(* IEC 61131-3 sources: plc-st-coding-agent/progress/evidence/f14_v10_full_20261113/jobs/custom_deepseek-v4pro, 130 files *)

(* ---- public-easy-01.candidate_01.st ---- *)
(*
ENGINEERING_CONTRACT
- Pump_Motor: active in state Cleaning, set by bottleSensor true when idle, retained until cleaningConfirmButton true (PUB001-PUB003).
- Filling_Valve: active in state Filling, set by cleaningConfirmButton true in Cleaning, retained until fillingConfirmButton true (PUB003-PUB004).
- Capping_Machine: active in state Capping, set by fillingConfirmButton true in Filling, retained until cappingConfirmButton true (PUB004-PUB005).
- Packing_Machine: active in state Packing, set by cappingConfirmButton true in Capping, retained until packingConfirmButton true (PUB005-PUB006).
- Completion_Light: active in state Done, set by packingConfirmButton true in Packing, retained until finishedButton true (PUB006-PUB007).
- Same-scan priority: exactly one transition evaluated per scan via IF/ELSIF on current state; outputs updated after transition.
- Units/boundaries: all signals are BOOL; state is an integer constant 0..5; no timing or analog units involved.
*)
(* CONTRACT_RULES [] *)

FUNCTION_BLOCK AutomatedFillingLineControl
VAR CONSTANT
    ST_IDLE : INT := 0;
    ST_CLEANING : INT := 1;
    ST_FILLING : INT := 2;
    ST_CAPPING : INT := 3;
    ST_PACKING : INT := 4;
    ST_DONE : INT := 5;
END_VAR
VAR
    state : INT := 0; (* initial idle state *)
END_VAR

IF state = ST_IDLE THEN
    IF bottleSensor THEN
        state := ST_CLEANING;
    END_IF;
ELSIF state = ST_CLEANING THEN
    IF cleaningConfirmButton THEN
        state := ST_FILLING;
    END_IF;
ELSIF state = ST_FILLING THEN
    IF fillingConfirmButton THEN
        state := ST_CAPPING;
    END_IF;
ELSIF state = ST_CAPPING THEN
    IF cappingConfirmButton THEN
        state := ST_PACKING;
    END_IF;
ELSIF state = ST_PACKING THEN
    IF packingConfirmButton THEN
        state := ST_DONE;
    END_IF;
ELSIF state = ST_DONE THEN
    IF finishedButton THEN
        state := ST_IDLE;
    END_IF;
END_IF;

Pump_Motor := (state = ST_CLEANING);
Filling_Valve := (state = ST_FILLING);
Capping_Machine := (state = ST_CAPPING);
Packing_Machine := (state = ST_PACKING);
Completion_Light := (state = ST_DONE);

END_FUNCTION_BLOCK

(* ---- public-easy-01.candidate_02.st ---- *)
(*
ENGINEERING_CONTRACT
- Pump_Motor: active in state Cleaning, set by bottleSensor true when idle, retained until cleaningConfirmButton true (PUB001-PUB003).
- Filling_Valve: active in state Filling, set by cleaningConfirmButton true in Cleaning, retained until fillingConfirmButton true (PUB003-PUB004).
- Capping_Machine: active in state Capping, set by fillingConfirmButton true in Filling, retained until cappingConfirmButton true (PUB004-PUB005).
- Packing_Machine: active in state Packing, set by cappingConfirmButton true in Capping, retained until packingConfirmButton true (PUB005-PUB006).
- Completion_Light: active in state Done, set by packingConfirmButton true in Packing, retained until finishedButton true (PUB006-PUB007).
- Same-scan priority: exactly one transition evaluated per scan via IF/ELSIF on current state; outputs updated after transition.
- Units/boundaries: all signals are BOOL; state is an integer constant 0..5; no timing or analog units involved.
*)
(* CONTRACT_RULES [] *)

FUNCTION_BLOCK AutomatedFillingLineControl
VAR_INPUT
    bottleSensor : BOOL;
    cleaningConfirmButton : BOOL;
    fillingConfirmButton : BOOL;
    cappingConfirmButton : BOOL;
    packingConfirmButton : BOOL;
    finishedButton : BOOL;
END_VAR
VAR_OUTPUT
    Pump_Motor : BOOL;
    Filling_Valve : BOOL;
    Capping_Machine : BOOL;
    Packing_Machine : BOOL;
    Completion_Light : BOOL;
END_VAR
VAR CONSTANT
    ST_IDLE : INT := 0;
    ST_CLEANING : INT := 1;
    ST_FILLING : INT := 2;
    ST_CAPPING : INT := 3;
    ST_PACKING : INT := 4;
    ST_DONE : INT := 5;
END_VAR
VAR
    state : INT := 0; (* initial idle state *)
END_VAR

IF state = ST_IDLE THEN
    IF bottleSensor THEN
        state := ST_CLEANING;
    END_IF;
ELSIF state = ST_CLEANING THEN
    IF cleaningConfirmButton THEN
        state := ST_FILLING;
    END_IF;
ELSIF state = ST_FILLING THEN
    IF fillingConfirmButton THEN
        state := ST_CAPPING;
    END_IF;
ELSIF state = ST_CAPPING THEN
    IF cappingConfirmButton THEN
        state := ST_PACKING;
    END_IF;
ELSIF state = ST_PACKING THEN
    IF packingConfirmButton THEN
        state := ST_DONE;
    END_IF;
ELSIF state = ST_DONE THEN
    IF finishedButton THEN
        state := ST_IDLE;
    END_IF;
END_IF;

Pump_Motor := (state = ST_CLEANING);
Filling_Valve := (state = ST_FILLING);
Capping_Machine := (state = ST_CAPPING);
Packing_Machine := (state = ST_PACKING);
Completion_Light := (state = ST_DONE);

END_FUNCTION_BLOCK

(* ---- public-easy-01.raw_candidate_01.st ---- *)
(*
ENGINEERING_CONTRACT
- Pump_Motor: active in state Cleaning, set by bottleSensor true when idle, retained until cleaningConfirmButton true (PUB001-PUB003).
- Filling_Valve: active in state Filling, set by cleaningConfirmButton true in Cleaning, retained until fillingConfirmButton true (PUB003-PUB004).
- Capping_Machine: active in state Capping, set by fillingConfirmButton true in Filling, retained until cappingConfirmButton true (PUB004-PUB005).
- Packing_Machine: active in state Packing, set by cappingConfirmButton true in Capping, retained until packingConfirmButton true (PUB005-PUB006).
- Completion_Light: active in state Done, set by packingConfirmButton true in Packing, retained until finishedButton true (PUB006-PUB007).
- Same-scan priority: exactly one transition evaluated per scan via IF/ELSIF on current state; outputs updated after transition.
- Units/boundaries: all signals are BOOL; state is an integer constant 0..5; no timing or analog units involved.
*)
(* CONTRACT_RULES [] *)

FUNCTION_BLOCK AutomatedFillingLineControl
VAR CONSTANT
    ST_IDLE : INT := 0;
    ST_CLEANING : INT := 1;
    ST_FILLING : INT := 2;
    ST_CAPPING : INT := 3;
    ST_PACKING : INT := 4;
    ST_DONE : INT := 5;
END_VAR
VAR
    state : INT := 0; (* initial idle state *)
END_VAR

IF state = ST_IDLE THEN
    IF bottleSensor THEN
        state := ST_CLEANING;
    END_IF;
ELSIF state = ST_CLEANING THEN
    IF cleaningConfirmButton THEN
        state := ST_FILLING;
    END_IF;
ELSIF state = ST_FILLING THEN
    IF fillingConfirmButton THEN
        state := ST_CAPPING;
    END_IF;
ELSIF state = ST_CAPPING THEN
    IF cappingConfirmButton THEN
        state := ST_PACKING;
    END_IF;
ELSIF state = ST_PACKING THEN
    IF packingConfirmButton THEN
        state := ST_DONE;
    END_IF;
ELSIF state = ST_DONE THEN
    IF finishedButton THEN
        state := ST_IDLE;
    END_IF;
END_IF;

Pump_Motor := (state = ST_CLEANING);
Filling_Valve := (state = ST_FILLING);
Capping_Machine := (state = ST_CAPPING);
Packing_Machine := (state = ST_PACKING);
Completion_Light := (state = ST_DONE);

END_FUNCTION_BLOCK

(* ---- public-easy-01.raw_candidate_02.st ---- *)
(*
ENGINEERING_CONTRACT
- Pump_Motor: active in state Cleaning, set by bottleSensor true when idle, retained until cleaningConfirmButton true (PUB001-PUB003).
- Filling_Valve: active in state Filling, set by cleaningConfirmButton true in Cleaning, retained until fillingConfirmButton true (PUB003-PUB004).
- Capping_Machine: active in state Capping, set by fillingConfirmButton true in Filling, retained until cappingConfirmButton true (PUB004-PUB005).
- Packing_Machine: active in state Packing, set by cappingConfirmButton true in Capping, retained until packingConfirmButton true (PUB005-PUB006).
- Completion_Light: active in state Done, set by packingConfirmButton true in Packing, retained until finishedButton true (PUB006-PUB007).
- Same-scan priority: exactly one transition evaluated per scan via IF/ELSIF on current state; outputs updated after transition.
- Units/boundaries: all signals are BOOL; state is an integer constant 0..5; no timing or analog units involved.
*)
(* CONTRACT_RULES [] *)

FUNCTION_BLOCK AutomatedFillingLineControl
VAR_INPUT
    bottleSensor : BOOL;
    cleaningConfirmButton : BOOL;
    fillingConfirmButton : BOOL;
    cappingConfirmButton : BOOL;
    packingConfirmButton : BOOL;
    finishedButton : BOOL;
END_VAR
VAR_OUTPUT
    Pump_Motor : BOOL;
    Filling_Valve : BOOL;
    Capping_Machine : BOOL;
    Packing_Machine : BOOL;
    Completion_Light : BOOL;
END_VAR
VAR CONSTANT
    ST_IDLE : INT := 0;
    ST_CLEANING : INT := 1;
    ST_FILLING : INT := 2;
    ST_CAPPING : INT := 3;
    ST_PACKING : INT := 4;
    ST_DONE : INT := 5;
END_VAR
VAR
    state : INT := 0; (* initial idle state *)
END_VAR

IF state = ST_IDLE THEN
    IF bottleSensor THEN
        state := ST_CLEANING;
    END_IF;
ELSIF state = ST_CLEANING THEN
    IF cleaningConfirmButton THEN
        state := ST_FILLING;
    END_IF;
ELSIF state = ST_FILLING THEN
    IF fillingConfirmButton THEN
        state := ST_CAPPING;
    END_IF;
ELSIF state = ST_CAPPING THEN
    IF cappingConfirmButton THEN
        state := ST_PACKING;
    END_IF;
ELSIF state = ST_PACKING THEN
    IF packingConfirmButton THEN
        state := ST_DONE;
    END_IF;
ELSIF state = ST_DONE THEN
    IF finishedButton THEN
        state := ST_IDLE;
    END_IF;
END_IF;

Pump_Motor := (state = ST_CLEANING);
Filling_Valve := (state = ST_FILLING);
Capping_Machine := (state = ST_CAPPING);
Packing_Machine := (state = ST_PACKING);
Completion_Light := (state = ST_DONE);

END_FUNCTION_BLOCK

(* ---- public-easy-02.candidate_01.st ---- *)
(*
ENGINEERING_CONTRACT
Activation: On every call after first, edge outputs computed from value vs lastValue.
Retention/hold: No latched outputs; all outputs are recomputed each scan from current and previous DWORD.
Reset/deactivation: No explicit reset; first invocation sets baseline lastValue:=value and reports no edges.
Same-scan priority: value is captured at scan start into lastValue after output computation; simultaneous change detection only.
Units/boundaries: risingBits/fallingBits are 32-bit DWORD masks, counts 0..32 as USINT; PUB001.
*)
(* CONTRACT_RULES [] *)

FUNCTION_BLOCK FB
VAR_INPUT
    value : DWORD;
END_VAR
VAR_OUTPUT
    hasChanged : BOOL;
    hasRisingEdges : BOOL;
    risingBits : DWORD;
    noOfRisingBits : USINT;
    hasFallingEdges : BOOL;
    fallingBits : DWORD;
    noOfFallingBits : USINT;
END_VAR
VAR
    lastValue : DWORD := DWORD#0;
    initialized : BOOL := FALSE;
    tmp_bits : DWORD;
    tmp_count : USINT;
    tmp_i : USINT;
END_VAR

// On first call, initialize previous value and report no changes/edges.
IF NOT initialized THEN
    lastValue := value;
    initialized := TRUE;
    hasChanged := FALSE;
    hasRisingEdges := FALSE;
    risingBits := DWORD#0;
    noOfRisingBits := USINT#0;
    hasFallingEdges := FALSE;
    fallingBits := DWORD#0;
    noOfFallingBits := USINT#0;
    RETURN;
END_IF;

// Compute changes and edge masks.
hasChanged := (value <> lastValue);
risingBits := value AND (NOT lastValue);
fallingBits := lastValue AND (NOT value);
hasRisingEdges := (risingBits <> DWORD#0);
hasFallingEdges := (fallingBits <> DWORD#0);

// Count rising edge bits.
tmp_count := USINT#0;
tmp_bits := risingBits;
FOR tmp_i := USINT#0 TO USINT#31 DO
    IF (tmp_bits AND DWORD#1) <> DWORD#0 THEN
        tmp_count := tmp_count + USINT#1;
    END_IF;
    tmp_bits := SHR(tmp_bits, UINT#1);
END_FOR;
noOfRisingBits := tmp_count;

// Count falling edge bits.
tmp_count := USINT#0;
tmp_bits := fallingBits;
FOR tmp_i := USINT#0 TO USINT#31 DO
    IF (tmp_bits AND DWORD#1) <> DWORD#0 THEN
        tmp_count := tmp_count + USINT#1;
    END_IF;
    tmp_bits := SHR(tmp_bits, UINT#1);
END_FOR;
noOfFallingBits := tmp_count;

// Store current value for next cycle.
lastValue := value;

END_FUNCTION_BLOCK

(* ---- public-easy-02.candidate_02.st ---- *)
(*
ENGINEERING_CONTRACT
Activation: On every call including first, edge outputs computed from value versus lastValue; lastValue initializes to 0.
Retention/hold: No latched outputs; all outputs are recomputed each scan from current and previous DWORD.
Reset/deactivation: No explicit reset; first invocation compares against zero and reports rising edges for set input bits.
Same-scan priority: value is captured before output computation; lastValue is updated at the end of the same invocation.
Units/boundaries: DWORD 32-bit masks, counts 0..32 as USINT; PUB001.
*)
(* CONTRACT_RULES [] *)

FUNCTION_BLOCK FB
VAR_INPUT
    value : DWORD;
END_VAR
VAR_OUTPUT
    hasChanged : BOOL;
    hasRisingEdges : BOOL;
    risingBits : DWORD;
    noOfRisingBits : USINT;
    hasFallingEdges : BOOL;
    fallingBits : DWORD;
    noOfFallingBits : USINT;
END_VAR
VAR
    lastValue : DWORD := DWORD#0;
    tmp_bits : DWORD;
    tmp_count : USINT;
    tmp_i : USINT;
END_VAR

hasChanged := (value <> lastValue);
risingBits := value AND (NOT lastValue);
fallingBits := lastValue AND (NOT value);
hasRisingEdges := (risingBits <> DWORD#0);
hasFallingEdges := (fallingBits <> DWORD#0);

tmp_count := USINT#0;
tmp_bits := risingBits;
FOR tmp_i := USINT#0 TO USINT#31 DO
    IF (tmp_bits AND DWORD#1) <> DWORD#0 THEN
        tmp_count := tmp_count + USINT#1;
    END_IF;
    tmp_bits := SHR(tmp_bits, UINT#1);
END_FOR;
noOfRisingBits := tmp_count;

tmp_count := USINT#0;
tmp_bits := fallingBits;
FOR tmp_i := USINT#0 TO USINT#31 DO
    IF (tmp_bits AND DWORD#1) <> DWORD#0 THEN
        tmp_count := tmp_count + USINT#1;
    END_IF;
    tmp_bits := SHR(tmp_bits, UINT#1);
END_FOR;
noOfFallingBits := tmp_count;

lastValue := value;

END_FUNCTION_BLOCK

(* ---- public-easy-02.raw_candidate_01.st ---- *)
(*
ENGINEERING_CONTRACT
Activation: On every call after first, edge outputs computed from value vs lastValue.
Retention/hold: No latched outputs; all outputs are recomputed each scan from current and previous DWORD.
Reset/deactivation: No explicit reset; first invocation sets baseline lastValue:=value and reports no edges.
Same-scan priority: value is captured at scan start into lastValue after output computation; simultaneous change detection only.
Units/boundaries: risingBits/fallingBits are 32-bit DWORD masks, counts 0..32 as USINT; PUB001.
*)
(* CONTRACT_RULES [] *)

FUNCTION_BLOCK FB
VAR_INPUT
    value : DWORD;
END_VAR
VAR_OUTPUT
    hasChanged : BOOL;
    hasRisingEdges : BOOL;
    risingBits : DWORD;
    noOfRisingBits : USINT;
    hasFallingEdges : BOOL;
    fallingBits : DWORD;
    noOfFallingBits : USINT;
END_VAR
VAR
    lastValue : DWORD := DWORD#0;
    initialized : BOOL := FALSE;
    tmp_bits : DWORD;
    tmp_count : USINT;
    tmp_i : USINT;
END_VAR

// On first call, initialize previous value and report no changes/edges.
IF NOT initialized THEN
    lastValue := value;
    initialized := TRUE;
    hasChanged := FALSE;
    hasRisingEdges := FALSE;
    risingBits := DWORD#0;
    noOfRisingBits := USINT#0;
    hasFallingEdges := FALSE;
    fallingBits := DWORD#0;
    noOfFallingBits := USINT#0;
    RETURN;
END_IF;

// Compute changes and edge masks.
hasChanged := (value <> lastValue);
risingBits := value AND (NOT lastValue);
fallingBits := lastValue AND (NOT value);
hasRisingEdges := (risingBits <> DWORD#0);
hasFallingEdges := (fallingBits <> DWORD#0);

// Count rising edge bits.
tmp_count := USINT#0;
tmp_bits := risingBits;
FOR tmp_i := USINT#0 TO USINT#31 DO
    IF (tmp_bits AND DWORD#1) <> DWORD#0 THEN
        tmp_count := tmp_count + USINT#1;
    END_IF;
    tmp_bits := SHR(tmp_bits, UINT#1);
END_FOR;
noOfRisingBits := tmp_count;

// Count falling edge bits.
tmp_count := USINT#0;
tmp_bits := fallingBits;
FOR tmp_i := USINT#0 TO USINT#31 DO
    IF (tmp_bits AND DWORD#1) <> DWORD#0 THEN
        tmp_count := tmp_count + USINT#1;
    END_IF;
    tmp_bits := SHR(tmp_bits, UINT#1);
END_FOR;
noOfFallingBits := tmp_count;

// Store current value for next cycle.
lastValue := value;

END_FUNCTION_BLOCK

(* ---- public-easy-02.raw_candidate_02.st ---- *)
(*
ENGINEERING_CONTRACT
Activation: On every call including first, edge outputs computed from value versus lastValue; lastValue initializes to 0.
Retention/hold: No latched outputs; all outputs are recomputed each scan from current and previous DWORD.
Reset/deactivation: No explicit reset; first invocation compares against zero and reports rising edges for set input bits.
Same-scan priority: value is captured before output computation; lastValue is updated at the end of the same invocation.
Units/boundaries: DWORD 32-bit masks, counts 0..32 as USINT; PUB001.
*)
(* CONTRACT_RULES [] *)

FUNCTION_BLOCK FB
VAR_INPUT
    value : DWORD;
END_VAR
VAR_OUTPUT
    hasChanged : BOOL;
    hasRisingEdges : BOOL;
    risingBits : DWORD;
    noOfRisingBits : USINT;
    hasFallingEdges : BOOL;
    fallingBits : DWORD;
    noOfFallingBits : USINT;
END_VAR
VAR
    lastValue : DWORD := DWORD#0;
    tmp_bits : DWORD;
    tmp_count : USINT;
    tmp_i : USINT;
END_VAR

hasChanged := (value <> lastValue);
risingBits := value AND (NOT lastValue);
fallingBits := lastValue AND (NOT value);
hasRisingEdges := (risingBits <> DWORD#0);
hasFallingEdges := (fallingBits <> DWORD#0);

tmp_count := USINT#0;
tmp_bits := risingBits;
FOR tmp_i := USINT#0 TO USINT#31 DO
    IF (tmp_bits AND DWORD#1) <> DWORD#0 THEN
        tmp_count := tmp_count + USINT#1;
    END_IF;
    tmp_bits := SHR(tmp_bits, UINT#1);
END_FOR;
noOfRisingBits := tmp_count;

tmp_count := USINT#0;
tmp_bits := fallingBits;
FOR tmp_i := USINT#0 TO USINT#31 DO
    IF (tmp_bits AND DWORD#1) <> DWORD#0 THEN
        tmp_count := tmp_count + USINT#1;
    END_IF;
    tmp_bits := SHR(tmp_bits, UINT#1);
END_FOR;
noOfFallingBits := tmp_count;

lastValue := value;

END_FUNCTION_BLOCK

(* ---- public-easy-03.candidate_01.st ---- *)
(* ENGINEERING_CONTRACT
   hiAlarm : SET on Value > hiLevel (PUB001), RESET on Value < hiLevel-hystWindow (PUB002), otherwise hold previous state.
   loAlarm : SET on Value < loLevel (PUB003), RESET on Value > loLevel+hystWindow (PUB004), otherwise hold previous state.
   error/status : SET 16#8001 when loLevel>=hiLevel and return (PUB005); SET 16#8002 when hystWindow>=hiLevel-loLevel and return (PUB006); cleared to FALSE/0 before checks.
   Priority : error checks run before alarm update; error returns preserve last alarm outputs.
   Boundaries : strict > and < for activation/deactivation; exact threshold equality holds current state. Negative hystWindow unspecified; applied as supplied.
   Units : REAL thresholds and values; status is WORD hex code.
*)
(* CONTRACT_RULES [] *)
FUNCTION_BLOCK AlarmHandling
VAR_INPUT
    Value : REAL;
    hiLevel : REAL;
    loLevel : REAL;
    hystWindow : REAL;
END_VAR
VAR_OUTPUT
    hiAlarm : BOOL;
    loAlarm : BOOL;
    error : BOOL;
    status : WORD;
END_VAR
VAR
END_VAR

    error := FALSE;
    status := 0;

    IF loLevel >= hiLevel THEN
        error := TRUE;
        status := 16#8001;
        RETURN;
    END_IF;

    IF hystWindow >= (hiLevel - loLevel) THEN
        error := TRUE;
        status := 16#8002;
        RETURN;
    END_IF;

    IF Value > hiLevel THEN
        hiAlarm := TRUE;
    ELSIF Value < (hiLevel - hystWindow) THEN
        hiAlarm := FALSE;
    END_IF;

    IF Value < loLevel THEN
        loAlarm := TRUE;
    ELSIF Value > (loLevel + hystWindow) THEN
        loAlarm := FALSE;
    END_IF;

END_FUNCTION_BLOCK

(* ---- public-easy-03.raw_candidate_01.st ---- *)
(* ENGINEERING_CONTRACT
   hiAlarm : SET on Value > hiLevel (PUB001), RESET on Value < hiLevel-hystWindow (PUB002), otherwise hold previous state.
   loAlarm : SET on Value < loLevel (PUB003), RESET on Value > loLevel+hystWindow (PUB004), otherwise hold previous state.
   error/status : SET 16#8001 when loLevel>=hiLevel and return (PUB005); SET 16#8002 when hystWindow>=hiLevel-loLevel and return (PUB006); cleared to FALSE/0 before checks.
   Priority : error checks run before alarm update; error returns preserve last alarm outputs.
   Boundaries : strict > and < for activation/deactivation; exact threshold equality holds current state. Negative hystWindow unspecified; applied as supplied.
   Units : REAL thresholds and values; status is WORD hex code.
*)
(* CONTRACT_RULES [] *)
FUNCTION_BLOCK AlarmHandling
VAR_INPUT
    Value : REAL;
    hiLevel : REAL;
    loLevel : REAL;
    hystWindow : REAL;
END_VAR
VAR_OUTPUT
    hiAlarm : BOOL;
    loAlarm : BOOL;
    error : BOOL;
    status : WORD;
END_VAR
VAR
END_VAR

    error := FALSE;
    status := 0;

    IF loLevel >= hiLevel THEN
        error := TRUE;
        status := 16#8001;
        RETURN;
    END_IF;

    IF hystWindow >= (hiLevel - loLevel) THEN
        error := TRUE;
        status := 16#8002;
        RETURN;
    END_IF;

    IF Value > hiLevel THEN
        hiAlarm := TRUE;
    ELSIF Value < (hiLevel - hystWindow) THEN
        hiAlarm := FALSE;
    END_IF;

    IF Value < loLevel THEN
        loAlarm := TRUE;
    ELSIF Value > (loLevel + hystWindow) THEN
        loAlarm := FALSE;
    END_IF;

END_FUNCTION_BLOCK

(* ---- public-easy-04.candidate_01.st ---- *)
(*
ENGINEERING_CONTRACT
1. DebounceValid state: set only while VISCOSITY_OK=TRUE and PASTE_E_STOP_NC=TRUE after accumulated CycleTime >= DebounceTime; immediate invalidation when VISCOSITY_OK=FALSE; incomplete timing is cleared when E-stop is FALSE (PUB001, PUB002).
2. VFD_RUN: active = PASTE_E_STOP_NC AND DebounceValid; E-stop has immediate priority and disables output in the same scan; no output latching (PUB002).
3. PUMP_RUNTIME_ACC: accumulates TO_LTIME(CycleTime) only when same-scan VFD_RUN=TRUE; preserves accumulated time while stopped; initial value 0 (PUB003, PUB005).
4. PUMP_MAINT_DUE: set when PUMP_RUNTIME_ACC >= LTIME#500H; because runtime is monotonic, it remains set; informational only with no effect on run/permissive logic (PUB004).
5. Initialization: VFD_RUN=FALSE, PUMP_RUNTIME_ACC=LTIME#0S, PUMP_MAINT_DUE=FALSE via declared initial values (PUB005).
Boundary: threshold comparisons use >= and TIME values are converted to LTIME; first satisfying debounce tick occurs when accumulated CycleTime reaches DebounceTime.
Unspecified: non-positive DebounceTime or CycleTime are assumed to be supplied positive (PUB006).
*)
(* CONTRACT_RULES [] *)
FUNCTION_BLOCK JamPump
VAR_INPUT
    VISCOSITY_OK : BOOL;
    PASTE_E_STOP_NC : BOOL;
    DebounceTime : TIME;
    CycleTime : TIME;
END_VAR
VAR_OUTPUT
    VFD_RUN : BOOL := FALSE;
    PUMP_MAINT_DUE : BOOL := FALSE;
    PUMP_RUNTIME_ACC : LTIME := LTIME#0S;
END_VAR
VAR
    local_DebounceElapsed : LTIME := LTIME#0S;
    local_ViscCondValid : BOOL := FALSE;
    local_MaintenanceLimit : LTIME := LTIME#500H;
END_VAR

IF NOT VISCOSITY_OK THEN
    local_ViscCondValid := FALSE;
    local_DebounceElapsed := LTIME#0S;
ELSE
    IF NOT PASTE_E_STOP_NC THEN
        IF NOT local_ViscCondValid THEN
            local_DebounceElapsed := LTIME#0S;
        END_IF;
    ELSE
        IF NOT local_ViscCondValid THEN
            local_DebounceElapsed := local_DebounceElapsed + TO_LTIME(CycleTime);
            IF local_DebounceElapsed >= TO_LTIME(DebounceTime) THEN
                local_ViscCondValid := TRUE;
            END_IF;
        END_IF;
    END_IF;
END_IF;

VFD_RUN := PASTE_E_STOP_NC AND local_ViscCondValid;

IF VFD_RUN THEN
    PUMP_RUNTIME_ACC := PUMP_RUNTIME_ACC + TO_LTIME(CycleTime);
END_IF;

PUMP_MAINT_DUE := (PUMP_RUNTIME_ACC >= local_MaintenanceLimit);

END_FUNCTION_BLOCK

(* ---- public-easy-04.raw_candidate_01.st ---- *)
(*
ENGINEERING_CONTRACT
1. DebounceValid state: set only while VISCOSITY_OK=TRUE and PASTE_E_STOP_NC=TRUE after accumulated CycleTime >= DebounceTime; immediate invalidation when VISCOSITY_OK=FALSE; incomplete timing is cleared when E-stop is FALSE (PUB001, PUB002).
2. VFD_RUN: active = PASTE_E_STOP_NC AND DebounceValid; E-stop has immediate priority and disables output in the same scan; no output latching (PUB002).
3. PUMP_RUNTIME_ACC: accumulates TO_LTIME(CycleTime) only when same-scan VFD_RUN=TRUE; preserves accumulated time while stopped; initial value 0 (PUB003, PUB005).
4. PUMP_MAINT_DUE: set when PUMP_RUNTIME_ACC >= LTIME#500H; because runtime is monotonic, it remains set; informational only with no effect on run/permissive logic (PUB004).
5. Initialization: VFD_RUN=FALSE, PUMP_RUNTIME_ACC=LTIME#0S, PUMP_MAINT_DUE=FALSE via declared initial values (PUB005).
Boundary: threshold comparisons use >= and TIME values are converted to LTIME; first satisfying debounce tick occurs when accumulated CycleTime reaches DebounceTime.
Unspecified: non-positive DebounceTime or CycleTime are assumed to be supplied positive (PUB006).
*)
(* CONTRACT_RULES [] *)
FUNCTION_BLOCK JamPump
VAR_INPUT
    VISCOSITY_OK : BOOL;
    PASTE_E_STOP_NC : BOOL;
    DebounceTime : TIME;
    CycleTime : TIME;
END_VAR
VAR_OUTPUT
    VFD_RUN : BOOL := FALSE;
    PUMP_MAINT_DUE : BOOL := FALSE;
    PUMP_RUNTIME_ACC : LTIME := LTIME#0S;
END_VAR
VAR
    local_DebounceElapsed : LTIME := LTIME#0S;
    local_ViscCondValid : BOOL := FALSE;
    local_MaintenanceLimit : LTIME := LTIME#500H;
END_VAR

IF NOT VISCOSITY_OK THEN
    local_ViscCondValid := FALSE;
    local_DebounceElapsed := LTIME#0S;
ELSE
    IF NOT PASTE_E_STOP_NC THEN
        IF NOT local_ViscCondValid THEN
            local_DebounceElapsed := LTIME#0S;
        END_IF;
    ELSE
        IF NOT local_ViscCondValid THEN
            local_DebounceElapsed := local_DebounceElapsed + TO_LTIME(CycleTime);
            IF local_DebounceElapsed >= TO_LTIME(DebounceTime) THEN
                local_ViscCondValid := TRUE;
            END_IF;
        END_IF;
    END_IF;
END_IF;

VFD_RUN := PASTE_E_STOP_NC AND local_ViscCondValid;

IF VFD_RUN THEN
    PUMP_RUNTIME_ACC := PUMP_RUNTIME_ACC + TO_LTIME(CycleTime);
END_IF;

PUMP_MAINT_DUE := (PUMP_RUNTIME_ACC >= local_MaintenanceLimit);

END_FUNCTION_BLOCK

(* ---- public-easy-05.candidate_01.st ---- *)
FUNCTION_BLOCK WeldGapAlarm
VAR_INPUT
    Gap_Exceeded: BOOL;
    Weld_E_Stop_NC: BOOL;
    DebounceTime: TIME;
END_VAR
VAR_OUTPUT
    Operator_Alert: BOOL;
    Weld_Soft_Start_Active: BOOL;
END_VAR
VAR
    tmp_InitTimer: TON;
    tmp_DebounceTimer: TON;
    local_InitActive: BOOL;
    local_EStopActive: BOOL;
    local_DebounceEnable: BOOL;
END_VAR

(* ENGINEERING_CONTRACT
   Output/Group         Activation                                      Retention/Hold                     Explicit Reset/Deactivation       Same-scan priority        Units/Bounds                  PUB
   Operator_Alert       Gap_Exceeded TRUE for DebounceTime after init   Holds while eligible gap TRUE      Gap FALSE, E-stop FALSE, init   E-stop overrides monitor   TIME, positive assumed        PUB003 PUB004
   Weld_Soft_Start_Act  5 s power-up init timer not elapsed             TRUE during init unless E-stop    E-stop active, timer elapsed     E-stop overrides init       TIME 5 s                      PUB002 PUB004 PUB005
   Debounce timing      eligible gap TRUE in normal monitoring         accumulates only if eligible       Gap FALSE, E-stop, init         E-stop/init clear timing    DebounceTime TIME             PUB002 PUB003 PUB004
*)

(* CONTRACT_RULES [] *)

local_EStopActive := NOT Weld_E_Stop_NC;

tmp_InitTimer(IN := TRUE, PT := T#5S);
local_InitActive := NOT tmp_InitTimer.Q;

local_DebounceEnable := Gap_Exceeded AND NOT local_InitActive AND NOT local_EStopActive;
tmp_DebounceTimer(IN := local_DebounceEnable, PT := DebounceTime);

Operator_Alert := tmp_DebounceTimer.Q AND NOT local_EStopActive;
Weld_Soft_Start_Active := local_InitActive AND NOT local_EStopActive;

END_FUNCTION_BLOCK

(* ---- public-easy-05.raw_candidate_01.st ---- *)
FUNCTION_BLOCK WeldGapAlarm
VAR_INPUT
    Gap_Exceeded: BOOL;
    Weld_E_Stop_NC: BOOL;
    DebounceTime: TIME;
END_VAR
VAR_OUTPUT
    Operator_Alert: BOOL;
    Weld_Soft_Start_Active: BOOL;
END_VAR
VAR
    tmp_InitTimer: TON;
    tmp_DebounceTimer: TON;
    local_InitActive: BOOL;
    local_EStopActive: BOOL;
    local_DebounceEnable: BOOL;
END_VAR

(* ENGINEERING_CONTRACT
   Output/Group         Activation                                      Retention/Hold                     Explicit Reset/Deactivation       Same-scan priority        Units/Bounds                  PUB
   Operator_Alert       Gap_Exceeded TRUE for DebounceTime after init   Holds while eligible gap TRUE      Gap FALSE, E-stop FALSE, init   E-stop overrides monitor   TIME, positive assumed        PUB003 PUB004
   Weld_Soft_Start_Act  5 s power-up init timer not elapsed             TRUE during init unless E-stop    E-stop active, timer elapsed     E-stop overrides init       TIME 5 s                      PUB002 PUB004 PUB005
   Debounce timing      eligible gap TRUE in normal monitoring         accumulates only if eligible       Gap FALSE, E-stop, init         E-stop/init clear timing    DebounceTime TIME             PUB002 PUB003 PUB004
*)

(* CONTRACT_RULES [] *)

local_EStopActive := NOT Weld_E_Stop_NC;

tmp_InitTimer(IN := TRUE, PT := T#5S);
local_InitActive := NOT tmp_InitTimer.Q;

local_DebounceEnable := Gap_Exceeded AND NOT local_InitActive AND NOT local_EStopActive;
tmp_DebounceTimer(IN := local_DebounceEnable, PT := DebounceTime);

Operator_Alert := tmp_DebounceTimer.Q AND NOT local_EStopActive;
Weld_Soft_Start_Active := local_InitActive AND NOT local_EStopActive;

END_FUNCTION_BLOCK

(* ---- public-easy-06.candidate_01.st ---- *)
FUNCTION_BLOCK AerationBlowerDelayedStart
VAR_INPUT
    DO_LOW : BOOL;
    AERATION_E_STOP_NC : BOOL;
END_VAR
VAR_OUTPUT
    BLOWER_RUN : BOOL := FALSE;
    AERATION_BLOWER_CYCLE_COUNT : UINT := 0;
END_VAR
VAR
    startTimer : TON;
    startEdge : R_TRIG;
END_VAR

(*
ENGINEERING_CONTRACT
Output BLOWER_RUN:
  activation: startTimer.Q after DO_LOW AND AERATION_E_STOP_NC true for T#5S (PUB001).
  hold: remains TRUE while both inputs stay TRUE (PUB001).
  reset/deactivation: DO_LOW=FALSE or AERATION_E_STOP_NC=FALSE disables same scan and resets timer (PUB002).
  units/boundaries: BOOL.
Output AERATION_BLOWER_CYCLE_COUNT:
  activation: increment on R_TRIG false->true of BLOWER_RUN (PUB003).
  hold: retains value during operation; stop does not reset count.
  reset: only power-up/cold init to 0 (PUB004).
  units/boundaries: UINT starts; saturates at 65535 (unspecified).
*)

(* CONTRACT_RULES [] *)

startTimer(IN := DO_LOW AND AERATION_E_STOP_NC, PT := T#5S);
BLOWER_RUN := startTimer.Q;

startEdge(CLK := BLOWER_RUN);
IF startEdge.Q THEN
    IF AERATION_BLOWER_CYCLE_COUNT < UINT#65535 THEN
        AERATION_BLOWER_CYCLE_COUNT := AERATION_BLOWER_CYCLE_COUNT + UINT#1;
    END_IF;
END_IF;

END_FUNCTION_BLOCK

(* ---- public-easy-06.raw_candidate_01.st ---- *)
FUNCTION_BLOCK AerationBlowerDelayedStart
VAR_INPUT
    DO_LOW : BOOL;
    AERATION_E_STOP_NC : BOOL;
END_VAR
VAR_OUTPUT
    BLOWER_RUN : BOOL := FALSE;
    AERATION_BLOWER_CYCLE_COUNT : UINT := 0;
END_VAR
VAR
    startTimer : TON;
    startEdge : R_TRIG;
END_VAR

(*
ENGINEERING_CONTRACT
Output BLOWER_RUN:
  activation: startTimer.Q after DO_LOW AND AERATION_E_STOP_NC true for T#5S (PUB001).
  hold: remains TRUE while both inputs stay TRUE (PUB001).
  reset/deactivation: DO_LOW=FALSE or AERATION_E_STOP_NC=FALSE disables same scan and resets timer (PUB002).
  units/boundaries: BOOL.
Output AERATION_BLOWER_CYCLE_COUNT:
  activation: increment on R_TRIG false->true of BLOWER_RUN (PUB003).
  hold: retains value during operation; stop does not reset count.
  reset: only power-up/cold init to 0 (PUB004).
  units/boundaries: UINT starts; saturates at 65535 (unspecified).
*)

(* CONTRACT_RULES [] *)

startTimer(IN := DO_LOW AND AERATION_E_STOP_NC, PT := T#5S);
BLOWER_RUN := startTimer.Q;

startEdge(CLK := BLOWER_RUN);
IF startEdge.Q THEN
    IF AERATION_BLOWER_CYCLE_COUNT < UINT#65535 THEN
        AERATION_BLOWER_CYCLE_COUNT := AERATION_BLOWER_CYCLE_COUNT + UINT#1;
    END_IF;
END_IF;

END_FUNCTION_BLOCK

(* ---- public-hard-01.candidate_01.st ---- *)
(* ENGINEERING_CONTRACT
   valveARun / valveBRun / valveCRun / valveDRun / mixMotorRun:
   - Activation: manual rising-edge toggle per PUB001; auto STATES OPEN_A/OPEN_B/WAIT_C/DONE/MIXING per PUB005-PUB010.
   - Retention: hold while selected mode/state condition remains; manual toggles hold until next edge, estop FALSE, or mode change.
   - Reset/deactivation: estop=FALSE forces all FALSE and resets manual/auto state; auto transitions close prior actuator; autoStart restart wins after transitions.
   - Same-scan priority: estop overrides all; manual outputs assigned only in manual; auto transitions selected on old state, then autoStart assignment wins.
   - levelSensor units cm, thresholds >=50, >=80, >=100; processMode sampled at 80 cm branch; mixMotorComplete edge accepted only while auto MIXING.
   - Unspecified: mode switch retains auto state; after estop clear, auto requires autoStart; manual requires button restart.
*)
(* CONTRACT_RULES [] *)

TYPE AUTO_STATE : (IDLE, OPEN_A, OPEN_B, WAIT_C, MIXING, DONE);
END_TYPE;

FUNCTION_BLOCK MaterialProportioningProcessControl
VAR_INPUT
    estop : BOOL;
    opeMode : BOOL;
    valveAStart : BOOL;
    valveBStart : BOOL;
    valveCStart : BOOL;
    valveDStart : BOOL;
    mixMotorStart : BOOL;
    autoStart : BOOL;
    processMode : BOOL;
    levelSensor : INT;
    mixMotorComplete : BOOL;
END_VAR
VAR_OUTPUT
    valveARun : BOOL;
    valveBRun : BOOL;
    valveCRun : BOOL;
    valveDRun : BOOL;
    mixMotorRun : BOOL;
END_VAR
VAR
    manualValveA : BOOL := FALSE;
    manualValveB : BOOL := FALSE;
    manualValveC : BOOL := FALSE;
    manualValveD : BOOL := FALSE;
    manualMixMotor : BOOL := FALSE;

    autoState : AUTO_STATE := AUTO_STATE#IDLE;

    rt_valveA : R_TRIG;
    rt_valveB : R_TRIG;
    rt_valveC : R_TRIG;
    rt_valveD : R_TRIG;
    rt_mixMotor : R_TRIG;
    rt_autoStart : R_TRIG;
    rt_mixComplete : R_TRIG;

    tmp_autoValveA : BOOL;
    tmp_autoValveB : BOOL;
    tmp_autoValveC : BOOL;
    tmp_autoValveD : BOOL;
    tmp_autoMixMotor : BOOL;
END_VAR

// Update rising-edge detectors
rt_valveA(CLK := valveAStart);
rt_valveB(CLK := valveBStart);
rt_valveC(CLK := valveCStart);
rt_valveD(CLK := valveDStart);
rt_mixMotor(CLK := mixMotorStart);
rt_autoStart(CLK := autoStart);
rt_mixComplete(CLK := mixMotorComplete);

// Emergency stop: reset all retained states while estop is FALSE
IF NOT estop THEN
    manualValveA := FALSE;
    manualValveB := FALSE;
    manualValveC := FALSE;
    manualValveD := FALSE;
    manualMixMotor := FALSE;
    autoState := AUTO_STATE#IDLE;
END_IF;

// Manual toggle controls only in manual mode with no emergency stop
IF estop AND NOT opeMode THEN
    IF rt_valveA.Q THEN
        manualValveA := NOT manualValveA;
    END_IF;
    IF rt_valveB.Q THEN
        manualValveB := NOT manualValveB;
    END_IF;
    IF rt_valveC.Q THEN
        manualValveC := NOT manualValveC;
    END_IF;
    IF rt_valveD.Q THEN
        manualValveD := NOT manualValveD;
    END_IF;
    IF rt_mixMotor.Q THEN
        manualMixMotor := NOT manualMixMotor;
    END_IF;
END_IF;

// Automatic process state transitions
IF estop AND opeMode THEN
    CASE autoState OF
        AUTO_STATE#OPEN_A:
            IF levelSensor >= 50 THEN
                autoState := AUTO_STATE#OPEN_B;
            END_IF;

        AUTO_STATE#OPEN_B:
            IF levelSensor >= 80 THEN
                IF NOT processMode THEN
                    autoState := AUTO_STATE#MIXING;
                ELSE
                    autoState := AUTO_STATE#WAIT_C;
                END_IF;
            END_IF;

        AUTO_STATE#WAIT_C:
            IF levelSensor >= 100 THEN
                autoState := AUTO_STATE#MIXING;
            END_IF;

        AUTO_STATE#MIXING:
            IF rt_mixComplete.Q THEN
                autoState := AUTO_STATE#DONE;
            END_IF;
    END_CASE;
END_IF;

// Auto start restarts the sequence and wins over same-scan state transitions
IF estop AND opeMode AND rt_autoStart.Q THEN
    autoState := AUTO_STATE#OPEN_A;
END_IF;

// Compute temporary automatic outputs from current state
tmp_autoValveA := FALSE;
tmp_autoValveB := FALSE;
tmp_autoValveC := FALSE;
tmp_autoValveD := FALSE;
tmp_autoMixMotor := FALSE;

CASE autoState OF
    AUTO_STATE#OPEN_A:
        tmp_autoValveA := TRUE;
    AUTO_STATE#OPEN_B:
        tmp_autoValveB := TRUE;
    AUTO_STATE#WAIT_C:
        tmp_autoValveC := TRUE;
    AUTO_STATE#MIXING:
        tmp_autoMixMotor := TRUE;
    AUTO_STATE#DONE:
        tmp_autoValveD := TRUE;
END_CASE;

// Final output assignment with emergency stop as highest priority
valveARun := FALSE;
valveBRun := FALSE;
valveCRun := FALSE;
valveDRun := FALSE;
mixMotorRun := FALSE;

IF estop AND NOT opeMode THEN
    valveARun := manualValveA;
    valveBRun := manualValveB;
    valveCRun := manualValveC;
    valveDRun := manualValveD;
    mixMotorRun := manualMixMotor;
ELSIF estop AND opeMode THEN
    valveARun := tmp_autoValveA;
    valveBRun := tmp_autoValveB;
    valveCRun := tmp_autoValveC;
    valveDRun := tmp_autoValveD;
    mixMotorRun := tmp_autoMixMotor;
END_IF;

END_FUNCTION_BLOCK

(* ---- public-hard-01.candidate_02.st ---- *)
(* ENGINEERING_CONTRACT
   valveARun / valveBRun / valveCRun / valveDRun / mixMotorRun:
   - Activation: manual rising-edge toggle per PUB001; auto STATES OPEN_A/OPEN_B/WAIT_C/DONE/MIXING per PUB005-PUB010.
   - Retention: hold while selected mode/state condition remains; manual toggles hold until next edge, estop FALSE, or mode change.
   - Reset/deactivation: estop=FALSE forces all FALSE and resets manual/auto state; auto transitions close prior actuator; autoStart restart wins after transitions.
   - Same-scan priority: estop overrides all; manual outputs assigned only in manual; auto transitions selected on old state, then autoStart assignment wins.
   - levelSensor units cm, thresholds >=50, >=80, >=100; processMode sampled at 80 cm branch; mixMotorComplete edge accepted only while auto MIXING.
   - Unspecified: mode switch retains auto state; after estop clear, auto requires autoStart; manual requires button restart.
*)
(* CONTRACT_RULES [] *)

TYPE AUTO_STATE : (IDLE, OPEN_A, OPEN_B, WAIT_C, MIXING, DONE);
END_TYPE;

FUNCTION_BLOCK MaterialProportioningProcessControl
VAR_INPUT
    estop : BOOL;
    opeMode : BOOL;
    valveAStart : BOOL;
    valveBStart : BOOL;
    valveCStart : BOOL;
    valveDStart : BOOL;
    mixMotorStart : BOOL;
    autoStart : BOOL;
    processMode : BOOL;
    levelSensor : INT;
    mixMotorComplete : BOOL;
END_VAR
VAR_OUTPUT
    valveARun : BOOL;
    valveBRun : BOOL;
    valveCRun : BOOL;
    valveDRun : BOOL;
    mixMotorRun : BOOL;
END_VAR
VAR
    manualValveA : BOOL := FALSE;
    manualValveB : BOOL := FALSE;
    manualValveC : BOOL := FALSE;
    manualValveD : BOOL := FALSE;
    manualMixMotor : BOOL := FALSE;

    autoState : AUTO_STATE := IDLE;

    rt_valveA : R_TRIG;
    rt_valveB : R_TRIG;
    rt_valveC : R_TRIG;
    rt_valveD : R_TRIG;
    rt_mixMotor : R_TRIG;
    rt_autoStart : R_TRIG;
    rt_mixComplete : R_TRIG;

    tmp_autoValveA : BOOL;
    tmp_autoValveB : BOOL;
    tmp_autoValveC : BOOL;
    tmp_autoValveD : BOOL;
    tmp_autoMixMotor : BOOL;
END_VAR

// Update rising-edge detectors
rt_valveA(CLK := valveAStart);
rt_valveB(CLK := valveBStart);
rt_valveC(CLK := valveCStart);
rt_valveD(CLK := valveDStart);
rt_mixMotor(CLK := mixMotorStart);
rt_autoStart(CLK := autoStart);
rt_mixComplete(CLK := mixMotorComplete);

// Emergency stop: reset all retained states while estop is FALSE
IF NOT estop THEN
    manualValveA := FALSE;
    manualValveB := FALSE;
    manualValveC := FALSE;
    manualValveD := FALSE;
    manualMixMotor := FALSE;
    autoState := IDLE;
END_IF;

// Manual toggle controls only in manual mode with no emergency stop
IF estop AND NOT opeMode THEN
    IF rt_valveA.Q THEN
        manualValveA := NOT manualValveA;
    END_IF;
    IF rt_valveB.Q THEN
        manualValveB := NOT manualValveB;
    END_IF;
    IF rt_valveC.Q THEN
        manualValveC := NOT manualValveC;
    END_IF;
    IF rt_valveD.Q THEN
        manualValveD := NOT manualValveD;
    END_IF;
    IF rt_mixMotor.Q THEN
        manualMixMotor := NOT manualMixMotor;
    END_IF;
END_IF;

// Automatic process state transitions
IF estop AND opeMode THEN
    CASE autoState OF
        OPEN_A:
            IF levelSensor >= 50 THEN
                autoState := OPEN_B;
            END_IF;

        OPEN_B:
            IF levelSensor >= 80 THEN
                IF NOT processMode THEN
                    autoState := MIXING;
                ELSE
                    autoState := WAIT_C;
                END_IF;
            END_IF;

        WAIT_C:
            IF levelSensor >= 100 THEN
                autoState := MIXING;
            END_IF;

        MIXING:
            IF rt_mixComplete.Q THEN
                autoState := DONE;
            END_IF;
    END_CASE;
END_IF;

// Auto start restarts the sequence and wins over same-scan state transitions
IF estop AND opeMode AND rt_autoStart.Q THEN
    autoState := OPEN_A;
END_IF;

// Compute temporary automatic outputs from current state
tmp_autoValveA := FALSE;
tmp_autoValveB := FALSE;
tmp_autoValveC := FALSE;
tmp_autoValveD := FALSE;
tmp_autoMixMotor := FALSE;

CASE autoState OF
    OPEN_A:
        tmp_autoValveA := TRUE;
    OPEN_B:
        tmp_autoValveB := TRUE;
    WAIT_C:
        tmp_autoValveC := TRUE;
    MIXING:
        tmp_autoMixMotor := TRUE;
    DONE:
        tmp_autoValveD := TRUE;
END_CASE;

// Final output assignment with emergency stop as highest priority
valveARun := FALSE;
valveBRun := FALSE;
valveCRun := FALSE;
valveDRun := FALSE;
mixMotorRun := FALSE;

IF estop AND NOT opeMode THEN
    valveARun := manualValveA;
    valveBRun := manualValveB;
    valveCRun := manualValveC;
    valveDRun := manualValveD;
    mixMotorRun := manualMixMotor;
ELSIF estop AND opeMode THEN
    valveARun := tmp_autoValveA;
    valveBRun := tmp_autoValveB;
    valveCRun := tmp_autoValveC;
    valveDRun := tmp_autoValveD;
    mixMotorRun := tmp_autoMixMotor;
END_IF;

END_FUNCTION_BLOCK

(* ---- public-hard-01.raw_candidate_01.st ---- *)
(* ENGINEERING_CONTRACT
   valveARun / valveBRun / valveCRun / valveDRun / mixMotorRun:
   - Activation: manual rising-edge toggle per PUB001; auto STATES OPEN_A/OPEN_B/WAIT_C/DONE/MIXING per PUB005-PUB010.
   - Retention: hold while selected mode/state condition remains; manual toggles hold until next edge, estop FALSE, or mode change.
   - Reset/deactivation: estop=FALSE forces all FALSE and resets manual/auto state; auto transitions close prior actuator; autoStart restart wins after transitions.
   - Same-scan priority: estop overrides all; manual outputs assigned only in manual; auto transitions selected on old state, then autoStart assignment wins.
   - levelSensor units cm, thresholds >=50, >=80, >=100; processMode sampled at 80 cm branch; mixMotorComplete edge accepted only while auto MIXING.
   - Unspecified: mode switch retains auto state; after estop clear, auto requires autoStart; manual requires button restart.
*)
(* CONTRACT_RULES [] *)

TYPE AUTO_STATE : (IDLE, OPEN_A, OPEN_B, WAIT_C, MIXING, DONE);
END_TYPE

FUNCTION_BLOCK MaterialProportioningProcessControl
VAR_INPUT
    estop : BOOL;
    opeMode : BOOL;
    valveAStart : BOOL;
    valveBStart : BOOL;
    valveCStart : BOOL;
    valveDStart : BOOL;
    mixMotorStart : BOOL;
    autoStart : BOOL;
    processMode : BOOL;
    levelSensor : INT;
    mixMotorComplete : BOOL;
END_VAR
VAR_OUTPUT
    valveARun : BOOL;
    valveBRun : BOOL;
    valveCRun : BOOL;
    valveDRun : BOOL;
    mixMotorRun : BOOL;
END_VAR
VAR
    manualValveA : BOOL := FALSE;
    manualValveB : BOOL := FALSE;
    manualValveC : BOOL := FALSE;
    manualValveD : BOOL := FALSE;
    manualMixMotor : BOOL := FALSE;

    autoState : AUTO_STATE := AUTO_STATE#IDLE;

    rt_valveA : R_TRIG;
    rt_valveB : R_TRIG;
    rt_valveC : R_TRIG;
    rt_valveD : R_TRIG;
    rt_mixMotor : R_TRIG;
    rt_autoStart : R_TRIG;
    rt_mixComplete : R_TRIG;

    tmp_autoValveA : BOOL;
    tmp_autoValveB : BOOL;
    tmp_autoValveC : BOOL;
    tmp_autoValveD : BOOL;
    tmp_autoMixMotor : BOOL;
END_VAR

// Update rising-edge detectors
rt_valveA(CLK := valveAStart);
rt_valveB(CLK := valveBStart);
rt_valveC(CLK := valveCStart);
rt_valveD(CLK := valveDStart);
rt_mixMotor(CLK := mixMotorStart);
rt_autoStart(CLK := autoStart);
rt_mixComplete(CLK := mixMotorComplete);

// Emergency stop: reset all retained states while estop is FALSE
IF NOT estop THEN
    manualValveA := FALSE;
    manualValveB := FALSE;
    manualValveC := FALSE;
    manualValveD := FALSE;
    manualMixMotor := FALSE;
    autoState := AUTO_STATE#IDLE;
END_IF

// Manual toggle controls only in manual mode with no emergency stop
IF estop AND NOT opeMode THEN
    IF rt_valveA.Q THEN
        manualValveA := NOT manualValveA;
    END_IF
    IF rt_valveB.Q THEN
        manualValveB := NOT manualValveB;
    END_IF
    IF rt_valveC.Q THEN
        manualValveC := NOT manualValveC;
    END_IF
    IF rt_valveD.Q THEN
        manualValveD := NOT manualValveD;
    END_IF
    IF rt_mixMotor.Q THEN
        manualMixMotor := NOT manualMixMotor;
    END_IF
END_IF

// Automatic process state transitions
IF estop AND opeMode THEN
    CASE autoState OF
        AUTO_STATE#OPEN_A:
            IF levelSensor >= 50 THEN
                autoState := AUTO_STATE#OPEN_B;
            END_IF

        AUTO_STATE#OPEN_B:
            IF levelSensor >= 80 THEN
                IF NOT processMode THEN
                    autoState := AUTO_STATE#MIXING;
                ELSE
                    autoState := AUTO_STATE#WAIT_C;
                END_IF
            END_IF

        AUTO_STATE#WAIT_C:
            IF levelSensor >= 100 THEN
                autoState := AUTO_STATE#MIXING;
            END_IF

        AUTO_STATE#MIXING:
            IF rt_mixComplete.Q THEN
                autoState := AUTO_STATE#DONE;
            END_IF
    END_CASE
END_IF

// Auto start restarts the sequence and wins over same-scan state transitions
IF estop AND opeMode AND rt_autoStart.Q THEN
    autoState := AUTO_STATE#OPEN_A;
END_IF

// Compute temporary automatic outputs from current state
tmp_autoValveA := FALSE;
tmp_autoValveB := FALSE;
tmp_autoValveC := FALSE;
tmp_autoValveD := FALSE;
tmp_autoMixMotor := FALSE;

CASE autoState OF
    AUTO_STATE#OPEN_A:
        tmp_autoValveA := TRUE;
    AUTO_STATE#OPEN_B:
        tmp_autoValveB := TRUE;
    AUTO_STATE#WAIT_C:
        tmp_autoValveC := TRUE;
    AUTO_STATE#MIXING:
        tmp_autoMixMotor := TRUE;
    AUTO_STATE#DONE:
        tmp_autoValveD := TRUE;
END_CASE

// Final output assignment with emergency stop as highest priority
valveARun := FALSE;
valveBRun := FALSE;
valveCRun := FALSE;
valveDRun := FALSE;
mixMotorRun := FALSE;

IF estop AND NOT opeMode THEN
    valveARun := manualValveA;
    valveBRun := manualValveB;
    valveCRun := manualValveC;
    valveDRun := manualValveD;
    mixMotorRun := manualMixMotor;
ELSIF estop AND opeMode THEN
    valveARun := tmp_autoValveA;
    valveBRun := tmp_autoValveB;
    valveCRun := tmp_autoValveC;
    valveDRun := tmp_autoValveD;
    mixMotorRun := tmp_autoMixMotor;
END_IF

END_FUNCTION_BLOCK

(* ---- public-hard-01.raw_candidate_02.st ---- *)
(* ENGINEERING_CONTRACT
   valveARun / valveBRun / valveCRun / valveDRun / mixMotorRun:
   - Activation: manual rising-edge toggle per PUB001; auto STATES OPEN_A/OPEN_B/WAIT_C/DONE/MIXING per PUB005-PUB010.
   - Retention: hold while selected mode/state condition remains; manual toggles hold until next edge, estop FALSE, or mode change.
   - Reset/deactivation: estop=FALSE forces all FALSE and resets manual/auto state; auto transitions close prior actuator; autoStart restart wins after transitions.
   - Same-scan priority: estop overrides all; manual outputs assigned only in manual; auto transitions selected on old state, then autoStart assignment wins.
   - levelSensor units cm, thresholds >=50, >=80, >=100; processMode sampled at 80 cm branch; mixMotorComplete edge accepted only while auto MIXING.
   - Unspecified: mode switch retains auto state; after estop clear, auto requires autoStart; manual requires button restart.
*)
(* CONTRACT_RULES [] *)

TYPE AUTO_STATE : (IDLE, OPEN_A, OPEN_B, WAIT_C, MIXING, DONE);
END_TYPE;

FUNCTION_BLOCK MaterialProportioningProcessControl
VAR_INPUT
    estop : BOOL;
    opeMode : BOOL;
    valveAStart : BOOL;
    valveBStart : BOOL;
    valveCStart : BOOL;
    valveDStart : BOOL;
    mixMotorStart : BOOL;
    autoStart : BOOL;
    processMode : BOOL;
    levelSensor : INT;
    mixMotorComplete : BOOL;
END_VAR
VAR_OUTPUT
    valveARun : BOOL;
    valveBRun : BOOL;
    valveCRun : BOOL;
    valveDRun : BOOL;
    mixMotorRun : BOOL;
END_VAR
VAR
    manualValveA : BOOL := FALSE;
    manualValveB : BOOL := FALSE;
    manualValveC : BOOL := FALSE;
    manualValveD : BOOL := FALSE;
    manualMixMotor : BOOL := FALSE;

    autoState : AUTO_STATE := IDLE;

    rt_valveA : R_TRIG;
    rt_valveB : R_TRIG;
    rt_valveC : R_TRIG;
    rt_valveD : R_TRIG;
    rt_mixMotor : R_TRIG;
    rt_autoStart : R_TRIG;
    rt_mixComplete : R_TRIG;

    tmp_autoValveA : BOOL;
    tmp_autoValveB : BOOL;
    tmp_autoValveC : BOOL;
    tmp_autoValveD : BOOL;
    tmp_autoMixMotor : BOOL;
END_VAR

// Update rising-edge detectors
rt_valveA(CLK := valveAStart);
rt_valveB(CLK := valveBStart);
rt_valveC(CLK := valveCStart);
rt_valveD(CLK := valveDStart);
rt_mixMotor(CLK := mixMotorStart);
rt_autoStart(CLK := autoStart);
rt_mixComplete(CLK := mixMotorComplete);

// Emergency stop: reset all retained states while estop is FALSE
IF NOT estop THEN
    manualValveA := FALSE;
    manualValveB := FALSE;
    manualValveC := FALSE;
    manualValveD := FALSE;
    manualMixMotor := FALSE;
    autoState := IDLE;
END_IF;

// Manual toggle controls only in manual mode with no emergency stop
IF estop AND NOT opeMode THEN
    IF rt_valveA.Q THEN
        manualValveA := NOT manualValveA;
    END_IF;
    IF rt_valveB.Q THEN
        manualValveB := NOT manualValveB;
    END_IF;
    IF rt_valveC.Q THEN
        manualValveC := NOT manualValveC;
    END_IF;
    IF rt_valveD.Q THEN
        manualValveD := NOT manualValveD;
    END_IF;
    IF rt_mixMotor.Q THEN
        manualMixMotor := NOT manualMixMotor;
    END_IF;
END_IF;

// Automatic process state transitions
IF estop AND opeMode THEN
    CASE autoState OF
        OPEN_A:
            IF levelSensor >= 50 THEN
                autoState := OPEN_B;
            END_IF;

        OPEN_B:
            IF levelSensor >= 80 THEN
                IF NOT processMode THEN
                    autoState := MIXING;
                ELSE
                    autoState := WAIT_C;
                END_IF;
            END_IF;

        WAIT_C:
            IF levelSensor >= 100 THEN
                autoState := MIXING;
            END_IF;

        MIXING:
            IF rt_mixComplete.Q THEN
                autoState := DONE;
            END_IF;
    END_CASE;
END_IF;

// Auto start restarts the sequence and wins over same-scan state transitions
IF estop AND opeMode AND rt_autoStart.Q THEN
    autoState := OPEN_A;
END_IF;

// Compute temporary automatic outputs from current state
tmp_autoValveA := FALSE;
tmp_autoValveB := FALSE;
tmp_autoValveC := FALSE;
tmp_autoValveD := FALSE;
tmp_autoMixMotor := FALSE;

CASE autoState OF
    OPEN_A:
        tmp_autoValveA := TRUE;
    OPEN_B:
        tmp_autoValveB := TRUE;
    WAIT_C:
        tmp_autoValveC := TRUE;
    MIXING:
        tmp_autoMixMotor := TRUE;
    DONE:
        tmp_autoValveD := TRUE;
END_CASE;

// Final output assignment with emergency stop as highest priority
valveARun := FALSE;
valveBRun := FALSE;
valveCRun := FALSE;
valveDRun := FALSE;
mixMotorRun := FALSE;

IF estop AND NOT opeMode THEN
    valveARun := manualValveA;
    valveBRun := manualValveB;
    valveCRun := manualValveC;
    valveDRun := manualValveD;
    mixMotorRun := manualMixMotor;
ELSIF estop AND opeMode THEN
    valveARun := tmp_autoValveA;
    valveBRun := tmp_autoValveB;
    valveCRun := tmp_autoValveC;
    valveDRun := tmp_autoValveD;
    mixMotorRun := tmp_autoMixMotor;
END_IF;

END_FUNCTION_BLOCK

(* ---- public-hard-02.candidate_01.st ---- *)
(* ENGINEERING_CONTRACT
- Outputs conveyorLeft/conveyorRight deactivate in IDLE, PROCESSING and DONE; active only in MOVING state; no latch. PUB005.
- State machine: 0=IDLE waits sensor1 AND station1Start with valid length; 1=MOVING waits arrival at target sensor; 2=PROCESSING waits completion at current station 2..4; 3=DONE after station 5 arrival. PUB001/PUB002/PUB005.
- Movement direction: target station > current -> conveyorRight; target < current -> conveyorLeft; target == current stays at station for repeated processing step. PUB005.
- Completion signals are level-sensitive; on receiving completion, step advances, next sequence entry is queried, and movement restarts toward that station. PUB002.
- Final active sequence entry is station 5; arrival at 5 stops conveyor and enters DONE. A new start is permitted from DONE when the start condition is true. PUB003/PUB006.
- processLength validated 1..8; dynamic array indexing bounded by processLength; sequence values assumed to satisfy contract (2..4 processing, final 5). PUB004.
- Unspecified: exact restart behavior after DONE is level-sensitive on sensor1 and station1Start. No explicit reset input is used.
*)
(* CONTRACT_RULES [] *)
FUNCTION_BLOCK FlexibleProcessingControl
VAR_INPUT
    processLength : USINT;
    sensor1 : BOOL;
    sensor2 : BOOL;
    sensor3 : BOOL;
    sensor4 : BOOL;
    sensor5 : BOOL;
    station1Start : BOOL;
    station2Complete : BOOL;
    station3Complete : BOOL;
    station4Complete : BOOL;
    processSequence : ARRAY[1..8] OF USINT;
END_VAR
VAR_OUTPUT
    conveyorLeft : BOOL;
    conveyorRight : BOOL;
END_VAR
VAR
    local_state : USINT := 0; (* 0 = idle, 1 = moving, 2 = processing, 3 = done *)
    local_step : USINT := 0;
    local_target : USINT := 0;
    local_currentStation : USINT := 1;
    local_moveLeft : BOOL := FALSE;
    local_moveRight : BOOL := FALSE;
    local_arrival : BOOL := FALSE;
    local_complete : BOOL := FALSE;
END_VAR

(* Default outputs deactivated unless set by MOVING state *)
conveyorLeft := FALSE;
conveyorRight := FALSE;

CASE local_state OF
0: (* IDLE: wait for raw material at station 1 and start button *)
    IF processLength >= 1 AND processLength <= 8 AND sensor1 AND station1Start THEN
        local_step := 1;
        local_target := processSequence[1];
        local_currentStation := 1;
        IF local_target > local_currentStation THEN
            local_moveLeft := FALSE;
            local_moveRight := TRUE;
            local_state := 1;
        ELSIF local_target < local_currentStation THEN
            local_moveLeft := TRUE;
            local_moveRight := FALSE;
            local_state := 1;
        ELSE
            (* target station 1 is outside the processing/output contract; remain idle *)
        END_IF;
    END_IF;

1: (* MOVING: drive conveyor in chosen direction until target sensor detects arrival *)
    conveyorLeft := local_moveLeft;
    conveyorRight := local_moveRight;

    local_arrival := FALSE;
    IF local_target = 1 AND sensor1 THEN
        local_arrival := TRUE;
    ELSIF local_target = 2 AND sensor2 THEN
        local_arrival := TRUE;
    ELSIF local_target = 3 AND sensor3 THEN
        local_arrival := TRUE;
    ELSIF local_target = 4 AND sensor4 THEN
        local_arrival := TRUE;
    ELSIF local_target = 5 AND sensor5 THEN
        local_arrival := TRUE;
    END_IF;

    IF local_arrival THEN
        conveyorLeft := FALSE;
        conveyorRight := FALSE;
        local_moveLeft := FALSE;
        local_moveRight := FALSE;
        local_currentStation := local_target;

        IF local_currentStation = 5 THEN
            local_state := 3; (* final output station reached *)
        ELSE
            local_state := 2; (* processing station reached *)
        END_IF;
    END_IF;

2: (* PROCESSING: wait for completion signal at current processing station *)
    local_complete := FALSE;
    IF local_currentStation = 2 THEN
        local_complete := station2Complete;
    ELSIF local_currentStation = 3 THEN
        local_complete := station3Complete;
    ELSIF local_currentStation = 4 THEN
        local_complete := station4Complete;
    END_IF;

    IF local_complete THEN
        IF local_step < processLength THEN
            local_step := local_step + 1;
            local_target := processSequence[local_step];

            IF local_target > local_currentStation THEN
                local_moveLeft := FALSE;
                local_moveRight := TRUE;
                local_state := 1;
            ELSIF local_target < local_currentStation THEN
                local_moveLeft := TRUE;
                local_moveRight := FALSE;
                local_state := 1;
            ELSE
                (* Same station: remain in processing for the next sequence entry *)
                local_state := 2;
            END_IF;
        ELSE
            (* Invalid sequence: current processing station is not followed by final station 5 *)
            local_state := 3;
        END_IF;
    END_IF;

3: (* DONE: product delivered to station 5; optionally wait for next start *)
    IF processLength >= 1 AND processLength <= 8 AND sensor1 AND station1Start THEN
        local_step := 1;
        local_target := processSequence[1];
        local_currentStation := 1;
        IF local_target > local_currentStation THEN
            local_moveLeft := FALSE;
            local_moveRight := TRUE;
            local_state := 1;
        ELSIF local_target < local_currentStation THEN
            local_moveLeft := TRUE;
            local_moveRight := FALSE;
            local_state := 1;
        ELSE
            (* target station 1 is outside the processing/output contract; remain done *)
        END_IF;
    END_IF;
END_CASE;

(* ---- public-hard-02.candidate_02.st ---- *)
(* ENGINEERING_CONTRACT
- Outputs conveyorLeft/deactivate in IDLE, PROCESSING and DONE; active only in MOVING state; no latch. PUB005.
- State machine: 0=IDLE waits sensor1 AND station1Start with valid length; 1=MOVING waits arrival at target sensor; 2=PROCESSING waits completion at current station 2..4; 3=DONE after station 5 arrival. PUB001/PUB002/PUB005.
- Movement direction: target station > current -> conveyorRight; target < current -> conveyorLeft; target == current stays at station for repeated processing step. PUB005.
- Completion signals are level-sensitive; on receiving completion, step advances, next sequence entry is queried, and movement restarts toward that station. PUB002.
- Final active sequence entry is station 5; arrival at 5 stops conveyor and enters DONE. A new start is permitted from DONE when the start condition is true. PUB003/PUB006.
- processLength validated 1..8; dynamic array indexing bounded by processLength; sequence values assumed to satisfy contract (2..4 processing, final 5). PUB004.
- Unspecified: exact restart behavior after DONE is level-sensitive on sensor1 and station1Start. No explicit reset input is used.
*)
(* CONTRACT_RULES [] *)
FUNCTION_BLOCK FlexibleProcessingControl
VAR_INPUT
    processLength : USINT;
    sensor1 : BOOL;
    sensor2 : BOOL;
    sensor3 : BOOL;
    sensor4 : BOOL;
    sensor5 : BOOL;
    station1Start : BOOL;
    station2Complete : BOOL;
    station3Complete : BOOL;
    station4Complete : BOOL;
    processSequence : ARRAY[1..8] OF USINT;
END_VAR
VAR_OUTPUT
    conveyorLeft : BOOL;
    conveyorRight : BOOL;
END_VAR
VAR
    local_state : USINT := 0; (* 0 = idle, 1 = moving, 2 = processing, 3 = done *)
    local_step : USINT := 0;
    local_target : USINT := 0;
    local_currentStation : USINT := 1;
    local_moveLeft : BOOL := FALSE;
    local_moveRight : BOOL := FALSE;
    local_arrival : BOOL := FALSE;
    local_complete : BOOL := FALSE;
END_VAR

(* Default outputs deactivated unless set by MOVING state *)
conveyorLeft := FALSE;
conveyorRight := FALSE;

CASE local_state OF
0: (* IDLE: wait for raw material at station 1 and start button *)
    IF processLength >= 1 AND processLength <= 8 AND sensor1 AND station1Start THEN
        local_step := 1;
        local_target := processSequence[1];
        local_currentStation := 1;
        IF local_target > local_currentStation THEN
            local_moveLeft := FALSE;
            local_moveRight := TRUE;
            local_state := 1;
        ELSIF local_target < local_currentStation THEN
            local_moveLeft := TRUE;
            local_moveRight := FALSE;
            local_state := 1;
        ELSE
            (* target station 1 is outside the processing/output contract; remain idle *)
        END_IF;
    END_IF;

1: (* MOVING: drive conveyor in chosen direction until target sensor detects arrival *)
    conveyorLeft := local_moveLeft;
    conveyorRight := local_moveRight;

    local_arrival := FALSE;
    IF local_target = 1 AND sensor1 THEN
        local_arrival := TRUE;
    ELSIF local_target = 2 AND sensor2 THEN
        local_arrival := TRUE;
    ELSIF local_target = 3 AND sensor3 THEN
        local_arrival := TRUE;
    ELSIF local_target = 4 AND sensor4 THEN
        local_arrival := TRUE;
    ELSIF local_target = 5 AND sensor5 THEN
        local_arrival := TRUE;
    END_IF;

    IF local_arrival THEN
        conveyorLeft := FALSE;
        conveyorRight := FALSE;
        local_moveLeft := FALSE;
        local_moveRight := FALSE;
        local_currentStation := local_target;

        IF local_currentStation = 5 THEN
            local_state := 3; (* final output station reached *)
        ELSE
            local_state := 2; (* processing station reached *)
        END_IF;
    END_IF;

2: (* PROCESSING: wait for completion signal at current processing station *)
    local_complete := FALSE;
    IF local_currentStation = 2 THEN
        local_complete := station2Complete;
    ELSIF local_currentStation = 3 THEN
        local_complete := station3Complete;
    ELSIF local_currentStation = 4 THEN
        local_complete := station4Complete;
    END_IF;

    IF local_complete THEN
        IF local_step < processLength THEN
            local_step := local_step + 1;
            local_target := processSequence[local_step];

            IF local_target > local_currentStation THEN
                local_moveLeft := FALSE;
                local_moveRight := TRUE;
                local_state := 1;
            ELSIF local_target < local_currentStation THEN
                local_moveLeft := TRUE;
                local_moveRight := FALSE;
                local_state := 1;
            ELSE
                (* Same station: remain in processing for the next sequence entry *)
                local_state := 2;
            END_IF;
        ELSE
            (* Invalid sequence: current processing station is not followed by final station 5 *)
            local_state := 3;
        END_IF;
    END_IF;

3: (* DONE: product delivered to station 5; optionally wait for next start *)
    IF processLength >= 1 AND processLength <= 8 AND sensor1 AND station1Start THEN
        local_step := 1;
        local_target := processSequence[1];
        local_currentStation := 1;
        IF local_target > local_currentStation THEN
            local_moveLeft := FALSE;
            local_moveRight := TRUE;
            local_state := 1;
        ELSIF local_target < local_currentStation THEN
            local_moveLeft := TRUE;
            local_moveRight := FALSE;
            local_state := 1;
        ELSE
            (* target station 1 is outside the processing/output contract; remain done *)
        END_IF;
    END_IF;
END_CASE;

END_FUNCTION_BLOCK

(* ---- public-hard-02.candidate_03.st ---- *)
(* ENGINEERING_CONTRACT
- Outputs conveyorLeft/deactivate in IDLE, PROCESSING and DONE; active only in MOVING state; no latch. PUB005.
- State machine: 0=IDLE waits sensor1 AND station1Start with valid length; 1=MOVING waits arrival at target sensor; 2=PROCESSING waits completion at current station 2..4; 3=DONE after station 5 arrival. PUB001/PUB002/PUB005.
- Movement direction: target station > current -> conveyorRight; target < current -> conveyorLeft; target == current stays at station for repeated processing step. PUB005.
- Completion signals are level-sensitive; on receiving completion, step advances, next sequence entry is queried, and movement restarts toward that station. PUB002.
- Final active sequence entry is station 5; arrival at 5 stops conveyor and enters DONE. A new start is permitted from DONE when the start condition is true. PUB003/PUB006.
- processLength validated 1..8; dynamic array indexing bounded by processLength; sequence values assumed to satisfy contract (2..4 processing, final 5). PUB004.
- Unspecified: exact restart behavior after DONE is level-sensitive on sensor1 and station1Start. No explicit reset input is used.
*)
(* CONTRACT_RULES [] *)
FUNCTION_BLOCK FlexibleProcessingControl
VAR_INPUT
    processLength : USINT;
    sensor1 : BOOL;
    sensor2 : BOOL;
    sensor3 : BOOL;
    sensor4 : BOOL;
    sensor5 : BOOL;
    station1Start : BOOL;
    station2Complete : BOOL;
    station3Complete : BOOL;
    station4Complete : BOOL;
    processSequence : ARRAY[1..8] OF USINT;
END_VAR
VAR_OUTPUT
    conveyorLeft : BOOL;
    conveyorRight : BOOL;
END_VAR
VAR
    local_state : USINT := 0; (* 0 = idle, 1 = moving, 2 = processing, 3 = done *)
    local_step : USINT := 0;
    local_target : USINT := 0;
    local_currentStation : USINT := 1;
    local_moveLeft : BOOL := FALSE;
    local_moveRight : BOOL := FALSE;
    local_arrival : BOOL := FALSE;
    local_complete : BOOL := FALSE;
END_VAR

(* Default outputs deactivated unless set by MOVING state *)
conveyorLeft := FALSE;
conveyorRight := FALSE;

CASE local_state OF
0: (* IDLE: wait for raw material at station 1 and start button *)
    IF processLength >= 1 AND processLength <= 8 AND sensor1 AND station1Start THEN
        local_step := 1;
        local_target := processSequence[1];
        local_currentStation := 1;
        IF local_target > local_currentStation THEN
            local_moveLeft := FALSE;
            local_moveRight := TRUE;
            local_state := 1;
        ELSIF local_target < local_currentStation THEN
            local_moveLeft := TRUE;
            local_moveRight := FALSE;
            local_state := 1;
        END_IF;
    END_IF;

1: (* MOVING: drive conveyor in chosen direction until target sensor detects arrival *)
    conveyorLeft := local_moveLeft;
    conveyorRight := local_moveRight;

    local_arrival := FALSE;
    IF local_target = 1 AND sensor1 THEN
        local_arrival := TRUE;
    ELSIF local_target = 2 AND sensor2 THEN
        local_arrival := TRUE;
    ELSIF local_target = 3 AND sensor3 THEN
        local_arrival := TRUE;
    ELSIF local_target = 4 AND sensor4 THEN
        local_arrival := TRUE;
    ELSIF local_target = 5 AND sensor5 THEN
        local_arrival := TRUE;
    END_IF;

    IF local_arrival THEN
        conveyorLeft := FALSE;
        conveyorRight := FALSE;
        local_moveLeft := FALSE;
        local_moveRight := FALSE;
        local_currentStation := local_target;

        IF local_currentStation = 5 THEN
            local_state := 3; (* final output station reached *)
        ELSE
            local_state := 2; (* processing station reached *)
        END_IF;
    END_IF;

2: (* PROCESSING: wait for completion signal at current processing station *)
    local_complete := FALSE;
    IF local_currentStation = 2 THEN
        local_complete := station2Complete;
    ELSIF local_currentStation = 3 THEN
        local_complete := station3Complete;
    ELSIF local_currentStation = 4 THEN
        local_complete := station4Complete;
    END_IF;

    IF local_complete THEN
        IF local_step < processLength THEN
            local_step := local_step + 1;
            local_target := processSequence[local_step];

            IF local_target > local_currentStation THEN
                local_moveLeft := FALSE;
                local_moveRight := TRUE;
                local_state := 1;
            ELSIF local_target < local_currentStation THEN
                local_moveLeft := TRUE;
                local_moveRight := FALSE;
                local_state := 1;
            ELSE
                (* Same station: remain in processing for the next sequence entry *)
                local_state := 2;
            END_IF;
        ELSE
            (* Invalid sequence: current processing station is not followed by final station 5 *)
            local_state := 3;
        END_IF;
    END_IF;

3: (* DONE: product delivered to station 5; optionally wait for next start *)
    IF processLength >= 1 AND processLength <= 8 AND sensor1 AND station1Start THEN
        local_step := 1;
        local_target := processSequence[1];
        local_currentStation := 1;
        IF local_target > local_currentStation THEN
            local_moveLeft := FALSE;
            local_moveRight := TRUE;
            local_state := 1;
        ELSIF local_target < local_currentStation THEN
            local_moveLeft := TRUE;
            local_moveRight := FALSE;
            local_state := 1;
        END_IF;
    END_IF;
END_CASE;

END_FUNCTION_BLOCK

(* ---- public-hard-02.candidate_04.st ---- *)
(* ENGINEERING_CONTRACT
- Outputs conveyorLeft/deactivate in IDLE, PROCESSING and DONE; active only in MOVING state; no latch. PUB005.
- State machine: 0=IDLE waits sensor1 AND station1Start with valid length; 1=MOVING waits arrival at target sensor; 2=PROCESSING waits completion at current station 2..4; 3=DONE after station 5 arrival. PUB001/PUB002/PUB005.
- Movement direction: target station > current -> conveyorRight; target < current -> conveyorLeft; target == current stays at station for repeated processing step. PUB005.
- Completion signals are level-sensitive; on receiving completion, step advances, next sequence entry is queried, and movement restarts toward that station. PUB002.
- Final active sequence entry is station 5; arrival at 5 stops conveyor and enters DONE. A new start is permitted from DONE when the start condition is true. PUB003/PUB006.
- processLength validated 1..8; dynamic array indexing bounded by processLength; sequence values assumed to satisfy contract (2..4 processing, final 5). PUB004.
- Unspecified: exact restart behavior after DONE is level-sensitive on sensor1 and station1Start. No explicit reset input is used.
*)
(* CONTRACT_RULES [] *)
FUNCTION_BLOCK FlexibleProcessingControl
VAR_INPUT
    processLength : USINT;
    sensor1 : BOOL;
    sensor2 : BOOL;
    sensor3 : BOOL;
    sensor4 : BOOL;
    sensor5 : BOOL;
    station1Start : BOOL;
    station2Complete : BOOL;
    station3Complete : BOOL;
    station4Complete : BOOL;
    processSequence : ARRAY[1..8] OF USINT;
END_VAR
VAR_OUTPUT
    conveyorLeft : BOOL;
    conveyorRight : BOOL;
END_VAR
VAR
    local_state : USINT := 0; (* 0 = idle, 1 = moving, 2 = processing, 3 = done *)
    local_step : USINT := 0;
    local_target : USINT := 0;
    local_currentStation : USINT := 1;
    local_moveLeft : BOOL := FALSE;
    local_moveRight : BOOL := FALSE;
    local_arrival : BOOL := FALSE;
    local_complete : BOOL := FALSE;
END_VAR

(* Default outputs deactivated unless set by MOVING state *)
conveyorLeft := FALSE;
conveyorRight := FALSE;

CASE local_state OF
0: (* IDLE: wait for raw material at station 1 and start button *)
    IF processLength >= 1 AND processLength <= 8 AND sensor1 AND station1Start THEN
        local_step := 1;
        local_target := processSequence[1];
        local_currentStation := 1;
        IF local_target > local_currentStation THEN
            local_moveLeft := FALSE;
            local_moveRight := TRUE;
            conveyorLeft := FALSE;
            conveyorRight := TRUE;
            local_state := 1;
        ELSIF local_target < local_currentStation THEN
            local_moveLeft := TRUE;
            local_moveRight := FALSE;
            conveyorLeft := TRUE;
            conveyorRight := FALSE;
            local_state := 1;
        END_IF;
    END_IF;

1: (* MOVING: drive conveyor in chosen direction until target sensor detects arrival *)
    conveyorLeft := local_moveLeft;
    conveyorRight := local_moveRight;

    local_arrival := FALSE;
    IF local_target = 1 AND sensor1 THEN
        local_arrival := TRUE;
    ELSIF local_target = 2 AND sensor2 THEN
        local_arrival := TRUE;
    ELSIF local_target = 3 AND sensor3 THEN
        local_arrival := TRUE;
    ELSIF local_target = 4 AND sensor4 THEN
        local_arrival := TRUE;
    ELSIF local_target = 5 AND sensor5 THEN
        local_arrival := TRUE;
    END_IF;

    IF local_arrival THEN
        conveyorLeft := FALSE;
        conveyorRight := FALSE;
        local_moveLeft := FALSE;
        local_moveRight := FALSE;
        local_currentStation := local_target;

        IF local_currentStation = 5 THEN
            local_state := 3; (* final output station reached *)
        ELSE
            local_state := 2; (* processing station reached *)
        END_IF;
    END_IF;

2: (* PROCESSING: wait for completion signal at current processing station *)
    local_complete := FALSE;
    IF local_currentStation = 2 THEN
        local_complete := station2Complete;
    ELSIF local_currentStation = 3 THEN
        local_complete := station3Complete;
    ELSIF local_currentStation = 4 THEN
        local_complete := station4Complete;
    END_IF;

    IF local_complete THEN
        IF local_step < processLength THEN
            local_step := local_step + 1;
            local_target := processSequence[local_step];

            IF local_target > local_currentStation THEN
                local_moveLeft := FALSE;
                local_moveRight := TRUE;
                conveyorLeft := FALSE;
                conveyorRight := TRUE;
                local_state := 1;
            ELSIF local_target < local_currentStation THEN
                local_moveLeft := TRUE;
                local_moveRight := FALSE;
                conveyorLeft := TRUE;
                conveyorRight := FALSE;
                local_state := 1;
            ELSE
                (* Same station: remain in processing for the next sequence entry *)
                local_state := 2;
            END_IF;
        ELSE
            (* Invalid sequence: current processing station is not followed by final station 5 *)
            local_state := 3;
        END_IF;
    END_IF;

3: (* DONE: product delivered to station 5; optionally wait for next start *)
    IF processLength >= 1 AND processLength <= 8 AND sensor1 AND station1Start THEN
        local_step := 1;
        local_target := processSequence[1];
        local_currentStation := 1;
        IF local_target > local_currentStation THEN
            local_moveLeft := FALSE;
            local_moveRight := TRUE;
            conveyorLeft := FALSE;
            conveyorRight := TRUE;
            local_state := 1;
        ELSIF local_target < local_currentStation THEN
            local_moveLeft := TRUE;
            local_moveRight := FALSE;
            conveyorLeft := TRUE;
            conveyorRight := FALSE;
            local_state := 1;
        END_IF;
    END_IF;
END_CASE;

END_FUNCTION_BLOCK

(* ---- public-hard-02.raw_candidate_01.st ---- *)
(* ENGINEERING_CONTRACT
- Outputs conveyorLeft/conveyorRight deactivate in IDLE, PROCESSING and DONE; active only in MOVING state; no latch. PUB005.
- State machine: 0=IDLE waits sensor1 AND station1Start with valid length; 1=MOVING waits arrival at target sensor; 2=PROCESSING waits completion at current station 2..4; 3=DONE after station 5 arrival. PUB001/PUB002/PUB005.
- Movement direction: target station > current -> conveyorRight; target < current -> conveyorLeft; target == current stays at station for repeated processing step. PUB005.
- Completion signals are level-sensitive; on receiving completion, step advances, next sequence entry is queried, and movement restarts toward that station. PUB002.
- Final active sequence entry is station 5; arrival at 5 stops conveyor and enters DONE. A new start is permitted from DONE when the start condition is true. PUB003/PUB006.
- processLength validated 1..8; dynamic array indexing bounded by processLength; sequence values assumed to satisfy contract (2..4 processing, final 5). PUB004.
- Unspecified: exact restart behavior after DONE is level-sensitive on sensor1 and station1Start. No explicit reset input is used.
*)
(* CONTRACT_RULES [] *)
FUNCTION_BLOCK FlexibleProcessingControl
VAR_INPUT
    processLength : USINT;
    sensor1 : BOOL;
    sensor2 : BOOL;
    sensor3 : BOOL;
    sensor4 : BOOL;
    sensor5 : BOOL;
    station1Start : BOOL;
    station2Complete : BOOL;
    station3Complete : BOOL;
    station4Complete : BOOL;
    processSequence : ARRAY[1..8] OF USINT;
END_VAR
VAR_OUTPUT
    conveyorLeft : BOOL;
    conveyorRight : BOOL;
END_VAR
VAR
    local_state : USINT := 0; (* 0 = idle, 1 = moving, 2 = processing, 3 = done *)
    local_step : USINT := 0;
    local_target : USINT := 0;
    local_currentStation : USINT := 1;
    local_moveLeft : BOOL := FALSE;
    local_moveRight : BOOL := FALSE;
    local_arrival : BOOL := FALSE;
    local_complete : BOOL := FALSE;
END_VAR

(* Default outputs deactivated unless set by MOVING state *)
conveyorLeft := FALSE;
conveyorRight := FALSE;

CASE local_state OF
0: (* IDLE: wait for raw material at station 1 and start button *)
    IF processLength >= 1 AND processLength <= 8 AND sensor1 AND station1Start THEN
        local_step := 1;
        local_target := processSequence[1];
        local_currentStation := 1;
        IF local_target > local_currentStation THEN
            local_moveLeft := FALSE;
            local_moveRight := TRUE;
            local_state := 1;
        ELSIF local_target < local_currentStation THEN
            local_moveLeft := TRUE;
            local_moveRight := FALSE;
            local_state := 1;
        ELSE
            (* target station 1 is outside the processing/output contract; remain idle *)
        END_IF;
    END_IF;

1: (* MOVING: drive conveyor in chosen direction until target sensor detects arrival *)
    conveyorLeft := local_moveLeft;
    conveyorRight := local_moveRight;

    local_arrival := FALSE;
    IF local_target = 1 AND sensor1 THEN
        local_arrival := TRUE;
    ELSIF local_target = 2 AND sensor2 THEN
        local_arrival := TRUE;
    ELSIF local_target = 3 AND sensor3 THEN
        local_arrival := TRUE;
    ELSIF local_target = 4 AND sensor4 THEN
        local_arrival := TRUE;
    ELSIF local_target = 5 AND sensor5 THEN
        local_arrival := TRUE;
    END_IF;

    IF local_arrival THEN
        conveyorLeft := FALSE;
        conveyorRight := FALSE;
        local_moveLeft := FALSE;
        local_moveRight := FALSE;
        local_currentStation := local_target;

        IF local_currentStation = 5 THEN
            local_state := 3; (* final output station reached *)
        ELSE
            local_state := 2; (* processing station reached *)
        END_IF;
    END_IF;

2: (* PROCESSING: wait for completion signal at current processing station *)
    local_complete := FALSE;
    IF local_currentStation = 2 THEN
        local_complete := station2Complete;
    ELSIF local_currentStation = 3 THEN
        local_complete := station3Complete;
    ELSIF local_currentStation = 4 THEN
        local_complete := station4Complete;
    END_IF;

    IF local_complete THEN
        IF local_step < processLength THEN
            local_step := local_step + 1;
            local_target := processSequence[local_step];

            IF local_target > local_currentStation THEN
                local_moveLeft := FALSE;
                local_moveRight := TRUE;
                local_state := 1;
            ELSIF local_target < local_currentStation THEN
                local_moveLeft := TRUE;
                local_moveRight := FALSE;
                local_state := 1;
            ELSE
                (* Same station: remain in processing for the next sequence entry *)
                local_state := 2;
            END_IF;
        ELSE
            (* Invalid sequence: current processing station is not followed by final station 5 *)
            local_state := 3;
        END_IF;
    END_IF;

3: (* DONE: product delivered to station 5; optionally wait for next start *)
    IF processLength >= 1 AND processLength <= 8 AND sensor1 AND station1Start THEN
        local_step := 1;
        local_target := processSequence[1];
        local_currentStation := 1;
        IF local_target > local_currentStation THEN
            local_moveLeft := FALSE;
            local_moveRight := TRUE;
            local_state := 1;
        ELSIF local_target < local_currentStation THEN
            local_moveLeft := TRUE;
            local_moveRight := FALSE;
            local_state := 1;
        ELSE
            (* target station 1 is outside the processing/output contract; remain done *)
        END_IF;
    END_IF;
END_CASE;

(* ---- public-hard-02.raw_candidate_02.st ---- *)
(* ENGINEERING_CONTRACT
- Outputs conveyorLeft/deactivate in IDLE, PROCESSING and DONE; active only in MOVING state; no latch. PUB005.
- State machine: 0=IDLE waits sensor1 AND station1Start with valid length; 1=MOVING waits arrival at target sensor; 2=PROCESSING waits completion at current station 2..4; 3=DONE after station 5 arrival. PUB001/PUB002/PUB005.
- Movement direction: target station > current -> conveyorRight; target < current -> conveyorLeft; target == current stays at station for repeated processing step. PUB005.
- Completion signals are level-sensitive; on receiving completion, step advances, next sequence entry is queried, and movement restarts toward that station. PUB002.
- Final active sequence entry is station 5; arrival at 5 stops conveyor and enters DONE. A new start is permitted from DONE when the start condition is true. PUB003/PUB006.
- processLength validated 1..8; dynamic array indexing bounded by processLength; sequence values assumed to satisfy contract (2..4 processing, final 5). PUB004.
- Unspecified: exact restart behavior after DONE is level-sensitive on sensor1 and station1Start. No explicit reset input is used.
*)
(* CONTRACT_RULES [] *)
FUNCTION_BLOCK FlexibleProcessingControl
VAR_INPUT
    processLength : USINT;
    sensor1 : BOOL;
    sensor2 : BOOL;
    sensor3 : BOOL;
    sensor4 : BOOL;
    sensor5 : BOOL;
    station1Start : BOOL;
    station2Complete : BOOL;
    station3Complete : BOOL;
    station4Complete : BOOL;
    processSequence : ARRAY[1..8] OF USINT;
END_VAR
VAR_OUTPUT
    conveyorLeft : BOOL;
    conveyorRight : BOOL;
END_VAR
VAR
    local_state : USINT := 0; (* 0 = idle, 1 = moving, 2 = processing, 3 = done *)
    local_step : USINT := 0;
    local_target : USINT := 0;
    local_currentStation : USINT := 1;
    local_moveLeft : BOOL := FALSE;
    local_moveRight : BOOL := FALSE;
    local_arrival : BOOL := FALSE;
    local_complete : BOOL := FALSE;
END_VAR

(* Default outputs deactivated unless set by MOVING state *)
conveyorLeft := FALSE;
conveyorRight := FALSE;

CASE local_state OF
0: (* IDLE: wait for raw material at station 1 and start button *)
    IF processLength >= 1 AND processLength <= 8 AND sensor1 AND station1Start THEN
        local_step := 1;
        local_target := processSequence[1];
        local_currentStation := 1;
        IF local_target > local_currentStation THEN
            local_moveLeft := FALSE;
            local_moveRight := TRUE;
            local_state := 1;
        ELSIF local_target < local_currentStation THEN
            local_moveLeft := TRUE;
            local_moveRight := FALSE;
            local_state := 1;
        ELSE
            (* target station 1 is outside the processing/output contract; remain idle *)
        END_IF;
    END_IF;

1: (* MOVING: drive conveyor in chosen direction until target sensor detects arrival *)
    conveyorLeft := local_moveLeft;
    conveyorRight := local_moveRight;

    local_arrival := FALSE;
    IF local_target = 1 AND sensor1 THEN
        local_arrival := TRUE;
    ELSIF local_target = 2 AND sensor2 THEN
        local_arrival := TRUE;
    ELSIF local_target = 3 AND sensor3 THEN
        local_arrival := TRUE;
    ELSIF local_target = 4 AND sensor4 THEN
        local_arrival := TRUE;
    ELSIF local_target = 5 AND sensor5 THEN
        local_arrival := TRUE;
    END_IF;

    IF local_arrival THEN
        conveyorLeft := FALSE;
        conveyorRight := FALSE;
        local_moveLeft := FALSE;
        local_moveRight := FALSE;
        local_currentStation := local_target;

        IF local_currentStation = 5 THEN
            local_state := 3; (* final output station reached *)
        ELSE
            local_state := 2; (* processing station reached *)
        END_IF;
    END_IF;

2: (* PROCESSING: wait for completion signal at current processing station *)
    local_complete := FALSE;
    IF local_currentStation = 2 THEN
        local_complete := station2Complete;
    ELSIF local_currentStation = 3 THEN
        local_complete := station3Complete;
    ELSIF local_currentStation = 4 THEN
        local_complete := station4Complete;
    END_IF;

    IF local_complete THEN
        IF local_step < processLength THEN
            local_step := local_step + 1;
            local_target := processSequence[local_step];

            IF local_target > local_currentStation THEN
                local_moveLeft := FALSE;
                local_moveRight := TRUE;
                local_state := 1;
            ELSIF local_target < local_currentStation THEN
                local_moveLeft := TRUE;
                local_moveRight := FALSE;
                local_state := 1;
            ELSE
                (* Same station: remain in processing for the next sequence entry *)
                local_state := 2;
            END_IF;
        ELSE
            (* Invalid sequence: current processing station is not followed by final station 5 *)
            local_state := 3;
        END_IF;
    END_IF;

3: (* DONE: product delivered to station 5; optionally wait for next start *)
    IF processLength >= 1 AND processLength <= 8 AND sensor1 AND station1Start THEN
        local_step := 1;
        local_target := processSequence[1];
        local_currentStation := 1;
        IF local_target > local_currentStation THEN
            local_moveLeft := FALSE;
            local_moveRight := TRUE;
            local_state := 1;
        ELSIF local_target < local_currentStation THEN
            local_moveLeft := TRUE;
            local_moveRight := FALSE;
            local_state := 1;
        ELSE
            (* target station 1 is outside the processing/output contract; remain done *)
        END_IF;
    END_IF;
END_CASE;

END_FUNCTION_BLOCK

(* ---- public-hard-02.raw_candidate_03.st ---- *)
(* ENGINEERING_CONTRACT
- Outputs conveyorLeft/deactivate in IDLE, PROCESSING and DONE; active only in MOVING state; no latch. PUB005.
- State machine: 0=IDLE waits sensor1 AND station1Start with valid length; 1=MOVING waits arrival at target sensor; 2=PROCESSING waits completion at current station 2..4; 3=DONE after station 5 arrival. PUB001/PUB002/PUB005.
- Movement direction: target station > current -> conveyorRight; target < current -> conveyorLeft; target == current stays at station for repeated processing step. PUB005.
- Completion signals are level-sensitive; on receiving completion, step advances, next sequence entry is queried, and movement restarts toward that station. PUB002.
- Final active sequence entry is station 5; arrival at 5 stops conveyor and enters DONE. A new start is permitted from DONE when the start condition is true. PUB003/PUB006.
- processLength validated 1..8; dynamic array indexing bounded by processLength; sequence values assumed to satisfy contract (2..4 processing, final 5). PUB004.
- Unspecified: exact restart behavior after DONE is level-sensitive on sensor1 and station1Start. No explicit reset input is used.
*)
(* CONTRACT_RULES [] *)
FUNCTION_BLOCK FlexibleProcessingControl
VAR_INPUT
    processLength : USINT;
    sensor1 : BOOL;
    sensor2 : BOOL;
    sensor3 : BOOL;
    sensor4 : BOOL;
    sensor5 : BOOL;
    station1Start : BOOL;
    station2Complete : BOOL;
    station3Complete : BOOL;
    station4Complete : BOOL;
    processSequence : ARRAY[1..8] OF USINT;
END_VAR
VAR_OUTPUT
    conveyorLeft : BOOL;
    conveyorRight : BOOL;
END_VAR
VAR
    local_state : USINT := 0; (* 0 = idle, 1 = moving, 2 = processing, 3 = done *)
    local_step : USINT := 0;
    local_target : USINT := 0;
    local_currentStation : USINT := 1;
    local_moveLeft : BOOL := FALSE;
    local_moveRight : BOOL := FALSE;
    local_arrival : BOOL := FALSE;
    local_complete : BOOL := FALSE;
END_VAR

(* Default outputs deactivated unless set by MOVING state *)
conveyorLeft := FALSE;
conveyorRight := FALSE;

CASE local_state OF
0: (* IDLE: wait for raw material at station 1 and start button *)
    IF processLength >= 1 AND processLength <= 8 AND sensor1 AND station1Start THEN
        local_step := 1;
        local_target := processSequence[1];
        local_currentStation := 1;
        IF local_target > local_currentStation THEN
            local_moveLeft := FALSE;
            local_moveRight := TRUE;
            local_state := 1;
        ELSIF local_target < local_currentStation THEN
            local_moveLeft := TRUE;
            local_moveRight := FALSE;
            local_state := 1;
        END_IF;
    END_IF;

1: (* MOVING: drive conveyor in chosen direction until target sensor detects arrival *)
    conveyorLeft := local_moveLeft;
    conveyorRight := local_moveRight;

    local_arrival := FALSE;
    IF local_target = 1 AND sensor1 THEN
        local_arrival := TRUE;
    ELSIF local_target = 2 AND sensor2 THEN
        local_arrival := TRUE;
    ELSIF local_target = 3 AND sensor3 THEN
        local_arrival := TRUE;
    ELSIF local_target = 4 AND sensor4 THEN
        local_arrival := TRUE;
    ELSIF local_target = 5 AND sensor5 THEN
        local_arrival := TRUE;
    END_IF;

    IF local_arrival THEN
        conveyorLeft := FALSE;
        conveyorRight := FALSE;
        local_moveLeft := FALSE;
        local_moveRight := FALSE;
        local_currentStation := local_target;

        IF local_currentStation = 5 THEN
            local_state := 3; (* final output station reached *)
        ELSE
            local_state := 2; (* processing station reached *)
        END_IF;
    END_IF;

2: (* PROCESSING: wait for completion signal at current processing station *)
    local_complete := FALSE;
    IF local_currentStation = 2 THEN
        local_complete := station2Complete;
    ELSIF local_currentStation = 3 THEN
        local_complete := station3Complete;
    ELSIF local_currentStation = 4 THEN
        local_complete := station4Complete;
    END_IF;

    IF local_complete THEN
        IF local_step < processLength THEN
            local_step := local_step + 1;
            local_target := processSequence[local_step];

            IF local_target > local_currentStation THEN
                local_moveLeft := FALSE;
                local_moveRight := TRUE;
                local_state := 1;
            ELSIF local_target < local_currentStation THEN
                local_moveLeft := TRUE;
                local_moveRight := FALSE;
                local_state := 1;
            ELSE
                (* Same station: remain in processing for the next sequence entry *)
                local_state := 2;
            END_IF;
        ELSE
            (* Invalid sequence: current processing station is not followed by final station 5 *)
            local_state := 3;
        END_IF;
    END_IF;

3: (* DONE: product delivered to station 5; optionally wait for next start *)
    IF processLength >= 1 AND processLength <= 8 AND sensor1 AND station1Start THEN
        local_step := 1;
        local_target := processSequence[1];
        local_currentStation := 1;
        IF local_target > local_currentStation THEN
            local_moveLeft := FALSE;
            local_moveRight := TRUE;
            local_state := 1;
        ELSIF local_target < local_currentStation THEN
            local_moveLeft := TRUE;
            local_moveRight := FALSE;
            local_state := 1;
        END_IF;
    END_IF;
END_CASE;

END_FUNCTION_BLOCK
